(* IEC 61131-3 sources: PortalRobot/Portal_robot/Device/application (part 4) *)

(* ---- PLC_PRG.RunSafety.st ---- *)
METHOD PRIVATE RunSafety

// --- BEGIN IMPLEMENTATION ---

FOR uiTwin := 1 TO 2 DO
	axTwinSafetyBusy[uiTwin] := (GVL_TWO_PALLET.uiMode = 1) AND (GVL_TWO_PALLET.astStatus[uiTwin].xBusy
		OR (GVL_TWO_PALLET.astInput[uiTwin].xAxisBound AND NOT GVL_TWO_PALLET.astInput[uiTwin].xStandstill));
END_FOR;
FOR uiMachine := UINT#1 TO UINT#4 DO
	axButtonStationInput[uiMachine] := GVL_CELL_SAFETY_IO.axDoorUnlockButtonInput[uiMachine]
		OR ((GVL_CELL_SETTINGS.eTestEnvironment = E_CELL_TEST_ENVIRONMENT.SIMULATION)
			AND GVL_CELL_SAFETY_IO.axSimDoorUnlockButtonInput[uiMachine]);
	axButtonStationEmergencyStopInput[uiMachine] := GVL_CELL_SAFETY_IO.axEmergencyStopButtonStationInput[uiMachine]
		OR ((GVL_CELL_SETTINGS.eTestEnvironment = E_CELL_TEST_ENVIRONMENT.SIMULATION)
			AND GVL_CELL_SAFETY_IO.axSimEmergencyStopButtonStationInput[uiMachine]);
END_FOR;
CELL_SAFETY(
	axMagazineMechanismBusy := axTwinSafetyBusy,
	axDoorLockClosedInput := GVL_CELL_SAFETY_IO.axDoorLockClosedInput,
	axDoorUnlockButtonInput := axButtonStationInput,
	axEmergencyStopButtonStationInput := axButtonStationEmergencyStopInput,
	axEmergencyStopCabinetInput := GVL_CELL_SAFETY_IO.axEmergencyStopCabinetInput,
	xEmergencyStopMpgInput := GVL_CELL_SAFETY_IO.xEmergencyStopMpgInput,
	xPhaseRelayOkInput := GVL_CELL_SAFETY_IO.xPhaseRelayOkInput,
	xPressureRelayOkInput := GVL_CELL_SAFETY_IO.xPressureRelayOkInput,
	xSafetyRelayOkInput := GVL_CELL_SAFETY_IO.xSafetyRelayOkInput,
	xCellStartButtonInput := GVL_CELL_SAFETY_IO.xCellStartButtonInput,
	xCellStopButtonInput := GVL_CELL_SAFETY_IO.xCellStopButtonInput,
	xCellResetButtonInput := GVL_CELL_SAFETY_IO.xCellResetButtonInput,
	xMpgAxisXInput := GVL_CELL_SAFETY_IO.xMpgAxisXInput,
	xMpgAxisYInput := GVL_CELL_SAFETY_IO.xMpgAxisYInput,
	xMpgAxisZInput := GVL_CELL_SAFETY_IO.xMpgAxisZInput,
	xMpgMultiplier1Input := GVL_CELL_SAFETY_IO.xMpgMultiplier1Input,
	xMpgMultiplier10Input := GVL_CELL_SAFETY_IO.xMpgMultiplier10Input,
	xMpgMultiplier100Input := GVL_CELL_SAFETY_IO.xMpgMultiplier100Input,
	xSafetyRelayReset := GVL_HMI.xSafetyRelayReset,
	astMagazineStatus := GVL_MAGAZINE.astStatus,
	FaultRequest := stSafetyFaultRequest
);

GVL_CELL_SAFETY_IO.axDoorUnlockOutput := CELL_SAFETY.axDoorUnlockOutput;
GVL_CELL_SAFETY_IO.axDoorButtonLampOutput := CELL_SAFETY.axDoorButtonLampOutput;
GVL_CELL_SAFETY_IO.xSafetyRelayResetOutput := CELL_SAFETY.xSafetyRelayResetOutput;

// Физические Старт/Стоп/Сброс — равноправные дубли HMI-команд, но только по фронту.
GVL_CELL_CONTROL.xEnable := GVL_CELL_CONTROL.xEnable OR CELL_SAFETY.xCellEnablePulse;
GVL_CELL_CONTROL.xDisable := GVL_CELL_CONTROL.xDisable OR CELL_SAFETY.xCellDisablePulse;
GVL_CELL_CONTROL.xReset := GVL_CELL_CONTROL.xReset OR CELL_SAFETY.xCellResetPulse;

// Ручное I/O владеет механизмами. Физический Start также не возобновляет
// прерванный автомат; выход из этого режима сам по себе ничего не запускает.
IF xIoManualActive THEN
	GVL_CELL_CONTROL.xStart := FALSE;
	GVL_CELL_CONTROL.xEnable := FALSE;
	GVL_CELL_CONTROL.xStop := TRUE;
END_IF;

CONTROLLER_DIAGNOSTICS(
    Request := GVL_HMI.stControllerWebRequest,
    udiNowMs := udiHmiCommandNowMs,
    xReset := GVL_CELL_CONTROL.xReset,
    xResetWarnings := GVL_ALARM.Command.xResetWarnings
);
GVL_HMI.stControllerWebStatus := CONTROLLER_DIAGNOSTICS.Status;
GVL_CELL_CONTROL.xGlobalError := CELL_SAFETY.Status.xGlobalError
    OR CONTROLLER_DIAGNOSTICS.Status.xGlobalStopRequired;
IF CONTROLLER_DIAGNOSTICS.Status.xAlarmActive THEN
    // Аппаратная системная авария не допускает обход через прямые ручные DO.
    xIoManualActive := FALSE;
    // Подтверждённое исчезновение причины разрешает восстановление, но не Auto.
    GVL_CELL_CONTROL.xStart := FALSE;
    GVL_CELL_CONTROL.xEnable := FALSE;
END_IF;

// HMI записывает payload, затем CommandSeq. Gateway удерживает единственного
// писателя до AckSeq. Даже запись между RunSafety и PublishHmi не теряется:
// PLC никогда не перезаписывает запрос, а обработает его в следующем скане.
uiCellModeRejectReason := UINT#0;
udiCellModeCommandSnapshot := GVL_HMI.udiCellModeCommandSeq;
IF (udiCellModeCommandSnapshot <> UDINT#0)
AND (udiCellModeCommandSnapshot <> GVL_HMI.udiCellModeAckSeq) THEN
	IF GVL_HMI.xCellManualRequest
	AND GVL_CELL_MANAGER.Status.xRunning
	AND NOT GVL_CELL_CONTROL.xGlobalError THEN
		uiCellModeRejectReason := UINT#2;
	ELSIF NOT GVL_HMI.xCellManualRequest
	AND (GVL_CELL_CONTROL.xGlobalError OR GVL_HMI.xIoEmergencyStopActive
        OR CONTROLLER_DIAGNOSTICS.Status.xAlarmActive) THEN
		uiCellModeRejectReason := UINT#3;
	ELSE
		GVL_CELL_CONTROL.xManual := GVL_HMI.xCellManualRequest;
	END_IF;
	IF uiCellModeRejectReason = UINT#0 THEN
		GVL_HMI.uiCellModeResult := UINT#1;
	ELSE
		GVL_HMI.uiCellModeResult := uiCellModeRejectReason;
	END_IF;
	// Ack публикуется после фактического режима в PublishHmi, включая отказ.
END_IF;

IF GVL_CELL_CONTROL.xGlobalError OR GVL_HMI.xIoEmergencyStopActive
OR CONTROLLER_DIAGNOSTICS.Status.xAlarmActive THEN
	GVL_CELL_CONTROL.xManual := TRUE;
END_IF;

// Разрешения рассчитываются после применения режима и Safety текущего скана.
xRobotHmiPermit := GVL_CELL_CONTROL.xManual AND NOT GVL_CELL_MANAGER.Status.xRunning
    AND NOT xIoManualActive
    AND NOT GVL_HMI.xIoEmergencyStopActive;
xRobotAutoPowerOff := NOT GVL_CELL_CONTROL.xManual
	AND (GVL_ROBOT.Status.xError
		OR GVL_AXIS.arrAxis[1].Status.xError
		OR GVL_AXIS.arrAxis[2].Status.xError
		OR GVL_AXIS.arrAxis[3].Status.xError
		OR GVL_AXIS_GROUP.AxisGroup.Status.xLocalError
		OR GVL_AXIS_GROUP.AxisGroup.Status.xLogicalError
		OR GVL_AXIS_GROUP.AxisGroup.Status.xGroupError);

(* ---- PLC_PRG.RunSignalTower.st ---- *)
METHOD PRIVATE RunSignalTower
VAR
	xBlink : BOOL;
END_VAR

// --- BEGIN IMPLEMENTATION ---

fbAlarmHorn(astSource := astAlarmSource, tDuration := GVL_CELL_SETTINGS.tAlarmHornDuration);
GVL_CELL_SAFETY_IO.xAlarmHornOutput := fbAlarmHorn.xSound;

// Приоритет: авария > предупреждение > работа > готовность > остановлена/не готова.
// Вызывать после RunAlarms: используются актуальные сводные состояния этого скана.
IF GVL_ALARM.Status.xAlarmActive THEN
	usiSignalTowerMode := USINT#4;
ELSIF GVL_ALARM.Status.xWarningActive THEN
	usiSignalTowerMode := USINT#3;
ELSIF GVL_CELL_MANAGER.Status.xRunning THEN
	usiSignalTowerMode := USINT#1;
ELSIF GVL_CELL_MANAGER.Status.xReadyToStart THEN
	usiSignalTowerMode := USINT#2;
ELSE
	usiSignalTowerMode := USINT#5;
END_IF;

xBlink := (usiSignalTowerMode = USINT#2) OR (usiSignalTowerMode = USINT#4);
tonSignalTowerBlink(
	IN := xBlink AND (usiSignalTowerMode = usiSignalTowerPreviousMode) AND NOT tonSignalTowerBlink.Q,
	PT := T#500MS
);
// Каждый новый режим начинается со включённой секции, без ожидания таймера.
IF (usiSignalTowerMode <> usiSignalTowerPreviousMode) OR NOT xBlink THEN
	xSignalTowerBlinkOn := TRUE;
ELSIF tonSignalTowerBlink.Q THEN
	xSignalTowerBlinkOn := NOT xSignalTowerBlinkOn;
END_IF;
usiSignalTowerPreviousMode := usiSignalTowerMode;

GVL_CELL_SAFETY_IO.xSignalTowerRedOutput := (usiSignalTowerMode = USINT#5)
	OR ((usiSignalTowerMode = USINT#4) AND xSignalTowerBlinkOn);
GVL_CELL_SAFETY_IO.xSignalTowerAmberOutput := usiSignalTowerMode = USINT#3;
GVL_CELL_SAFETY_IO.xSignalTowerGreenOutput := (usiSignalTowerMode = USINT#1)
	OR ((usiSignalTowerMode = USINT#2) AND xSignalTowerBlinkOn);

(* ---- PLC_PRG.RunStatistics.st ---- *)
METHOD PRIVATE RunStatistics

// --- BEGIN IMPLEMENTATION ---

STATISTIC_MAIN(
    xStart := GVL_CELL_MANAGER.Status.xRunning,
    uiSimulationTimeFactor := GVL_CELL_SETTINGS.uiSimulationTimeFactorApplied,
    eActiveAction := GVL_ROBOT.Diag.eActiveAction,
    eActivePoint := GVL_ROBOT.Diag.eActivePoint,
    xBusyMagazine := GVL_MAGAZINE.astStatus[1].xBusy OR GVL_MAGAZINE.astStatus[2].xBusy,
    xBusyMachine_1 := GVL_MACHINE.Status[1].xBusy,
    xBusyMachine_2 := GVL_MACHINE.Status[2].xBusy,
    xBusyMachine_3 := GVL_MACHINE.Status[3].xBusy,
    xCycleActiveMachine_1 := GVL_MACHINE.Status[1].stIo.xCycleActive,
    xCycleActiveMachine_2 := GVL_MACHINE.Status[2].stIo.xCycleActive,
    xCycleActiveMachine_3 := GVL_MACHINE.Status[3].stIo.xCycleActive,
    xBusyRobot := GVL_ROBOT.Status.xBusy,
    udiNowMs := TIME_TO_UDINT(TIME())
);

IF STATISTIC_MAIN.xUpdated THEN
    GVL_STATISTIC.stStatistic := STATISTIC_MAIN.stStatistic;
END_IF;

(* ---- PLC_PRG.RunTestControl.st ---- *)
METHOD PRIVATE RunTestControl

// --- BEGIN IMPLEMENTATION ---

// Test environment is independent from the robot control interface.
rtTestEnvironmentApply(CLK := GVL_HMI.xTestEnvironmentApply);
rtTestSpeedProfileApply(CLK := GVL_HMI.xTestSpeedProfileApply);
rtTestScenarioApply(CLK := GVL_HMI.xTestScenarioApply);
xTestInitializePulse := FALSE;
xTestAbortActive := GVL_HMI.xTestAbort
	AND GVL_HMI.xTestSessionActive
	AND (GVL_CELL_SETTINGS.eTestEnvironment = E_CELL_TEST_ENVIRONMENT.SIMULATION);

xTestStable := NOT GVL_CELL_MANAGER.Status.xRunning
	AND NOT GVL_ROBOT.Status.xBusy
	AND NOT GVL_MAGAZINE.astStatus[1].xBusy
	AND NOT GVL_MAGAZINE.astStatus[2].xBusy
	AND NOT GVL_TWO_PALLET.astStatus[1].xBusy
	AND NOT GVL_TWO_PALLET.astStatus[2].xBusy
	AND NOT GVL_GEOMETRY_CONTROL.astStatus[1].xDriveRunning
	AND NOT GVL_GEOMETRY_CONTROL.astStatus[2].xDriveRunning
	AND NOT GVL_GEOMETRY_CONTROL.astStatus[1].xResetBusy
	AND NOT GVL_GEOMETRY_CONTROL.astStatus[2].xResetBusy
	AND NOT GVL_GEOMETRY_CONTROL.astStatus[1].xReserved
	AND NOT GVL_GEOMETRY_CONTROL.astStatus[2].xReserved
	AND NOT xMotionBusy
	AND NOT SIMULATION_DYNAMICS.xBusy;
FOR uiTestIndex := UINT#1 TO UINT#3 DO
	xTestStable := xTestStable
		AND NOT GVL_MACHINE.Status[uiTestIndex].xBusy
		AND NOT GVL_MACHINE.Status[uiTestIndex].xProcessing;
END_FOR;

GVL_HMI.xTestEnvironmentChangeAllowed := xTestStable
	AND NOT GVL_TWO_PALLET.astInput[1].xPowered
	AND NOT GVL_TWO_PALLET.astInput[2].xPowered;
GVL_HMI.xTestScenarioApplyAllowed := xTestStable
	AND ((GVL_TWO_PALLET.uiMode = 0)
		OR ((GVL_TWO_PALLET.uiMode = 1)
			AND (GVL_CELL_SETTINGS.eTestEnvironment = E_CELL_TEST_ENVIRONMENT.SIMULATION)
			AND NOT GVL_HMI.xModbusMode
			AND GVL_TWO_PALLET.astStatus[1].xConfirmed
			AND GVL_TWO_PALLET.astStatus[2].xConfirmed
			AND (GVL_TWO_PALLET.astStatus[1].uiRobotPallet >= UINT#1)
			AND (GVL_TWO_PALLET.astStatus[1].uiRobotPallet <= UINT#2)
			AND (GVL_TWO_PALLET.astStatus[2].uiRobotPallet >= UINT#1)
			AND (GVL_TWO_PALLET.astStatus[2].uiRobotPallet <= UINT#2)
			AND GVL_TWO_PALLET.astInput[1].xStandstill
			AND GVL_TWO_PALLET.astInput[2].xStandstill))
	AND GVL_HMI.xTestSessionActive
	AND (GVL_CELL_SETTINGS.eTestEnvironment <> E_CELL_TEST_ENVIRONMENT.NORMAL)
	AND ((GVL_CELL_SETTINGS.eTestEnvironment <> E_CELL_TEST_ENVIRONMENT.SIMULATION)
		OR NOT GVL_ROBOT_MODBUS.xModeActive
		OR GVL_ROBOT_MODBUS.Status.xSimulatorActive);
// Старые OPC UA поля сохранены для совместимости; физический ключ исключён.
GVL_HMI.xSc500BenchKeyActive := FALSE;

IF rtTestEnvironmentApply.Q THEN
	GVL_HMI.uiTestRejectReason := UINT#0;
	IF NOT GVL_HMI.xTestEnvironmentChangeAllowed THEN
		GVL_HMI.uiTestRejectReason := UINT#1; // equipment is not idle
	ELSIF GVL_HMI.uiTestEnvironmentRequest > UINT#2 THEN
		GVL_HMI.uiTestRejectReason := UINT#2; // invalid environment
	ELSIF (GVL_HMI.uiTestEnvironmentRequest = UINT#2)
	AND NOT GVL_ROBOT_MODBUS.xModeActive THEN
		GVL_HMI.uiTestRejectReason := UINT#3; // bench requires Modbus
	ELSIF (GVL_HMI.uiTestEnvironmentRequest = UINT#1)
	AND GVL_ROBOT_MODBUS.xModeActive
	AND NOT GVL_ROBOT_MODBUS.Status.xSimulatorActive THEN
		GVL_HMI.uiTestRejectReason := UINT#4; // Python simulator marker missing
	ELSE
		CASE GVL_HMI.uiTestEnvironmentRequest OF
			UINT#0: GVL_CELL_SETTINGS.eTestEnvironment := E_CELL_TEST_ENVIRONMENT.NORMAL;
			UINT#1: GVL_CELL_SETTINGS.eTestEnvironment := E_CELL_TEST_ENVIRONMENT.SIMULATION;
			UINT#2: GVL_CELL_SETTINGS.eTestEnvironment := E_CELL_TEST_ENVIRONMENT.SC500_BENCH;
		END_CASE;
		IF GVL_CELL_SETTINGS.eTestEnvironment = E_CELL_TEST_ENVIRONMENT.NORMAL THEN
			GVL_CELL_SETTINGS.xErrorSimulationEnabled := FALSE;
		END_IF;
		GVL_CELL_SETTINGS.eTestSpeedProfile := E_TEST_SPEED_PROFILE.REALTIME;
	END_IF;
END_IF;

IF rtTestSpeedProfileApply.Q THEN
	GVL_HMI.uiTestRejectReason := UINT#0;
	IF (GVL_HMI.uiTestSpeedProfileRequest <= UINT#1)
	AND (GVL_CELL_SETTINGS.eTestEnvironment = E_CELL_TEST_ENVIRONMENT.SIMULATION) THEN
		IF GVL_HMI.uiTestSpeedProfileRequest = UINT#1 THEN
			GVL_CELL_SETTINGS.eTestSpeedProfile := E_TEST_SPEED_PROFILE.FAST;
			// В Modbus профиль по-прежнему владеет коэффициентом внешней модели.
			// В SoftMotion коэффициент задаёт ползунок, а применение выполняется
			// отдельной транзакцией только на границе следующего теста.
			IF GVL_ROBOT_MODBUS.xModeActive THEN
				GVL_CELL_SETTINGS.uiSimulationTimeFactor := UINT#250;
			END_IF;
		ELSE
			GVL_CELL_SETTINGS.eTestSpeedProfile := E_TEST_SPEED_PROFILE.REALTIME;
			IF GVL_ROBOT_MODBUS.xModeActive THEN
				GVL_CELL_SETTINGS.uiSimulationTimeFactor := UINT#1;
			END_IF;
		END_IF;
		GVL_HMI.uiSimulationTimeFactor := GVL_CELL_SETTINGS.uiSimulationTimeFactor;
	ELSE
		GVL_HMI.uiTestRejectReason := UINT#5; // speed profile is simulation-only
	END_IF;
END_IF;

IF rtTestScenarioApply.Q THEN
	GVL_HMI.uiTestScenarioResult := UINT#0;
	uiTestSlotCount := UINT#120;
	IF GVL_TWO_PALLET.uiMode = UINT#1 THEN uiTestSlotCount := UINT#96; END_IF;
	xTestScenarioValid := (GVL_HMI.stTestScenario.uiSchemaVersion = UINT#3)
		AND (GVL_HMI.stTestScenario.uiMagazineMode = GVL_TWO_PALLET.uiMode)
		AND (GVL_HMI.stTestScenario.udiLoadSeq <> UDINT#0)
		AND (GVL_HMI.stTestScenario.uiTypeCount >= UINT#1)
		AND (GVL_HMI.stTestScenario.uiTypeCount <= UINT#3);
	FOR uiTestIndex := UINT#1 TO UINT#3 DO
		xTestScenarioValid := xTestScenarioValid
			AND (GVL_HMI.stTestScenario.auiMachineState[uiTestIndex] <= UINT#3)
			AND (GVL_HMI.stTestScenario.auiMachineType[uiTestIndex] >= UINT#1)
			AND (GVL_HMI.stTestScenario.auiMachineType[uiTestIndex]
				<= GVL_HMI.stTestScenario.uiTypeCount);
	END_FOR;
	FOR uiTestIndex := UINT#1 TO uiTestSlotCount DO
		xTestScenarioValid := xTestScenarioValid
			AND (GVL_HMI.stTestScenario.auiSlotType[uiTestIndex] >= UINT#1)
			AND (GVL_HMI.stTestScenario.auiSlotType[uiTestIndex]
				<= GVL_HMI.stTestScenario.uiTypeCount);
		FOR uiTestMagazine := UINT#1 TO UINT#2 DO
			xTestScenarioValid := xTestScenarioValid
				AND (GVL_HMI.stTestScenario.aauiSlotContent[uiTestMagazine, uiTestIndex] <= UINT#2)
				AND (GVL_HMI.stTestScenario.aauiOperatorSlotContent[uiTestMagazine, uiTestIndex] <= UINT#2);
		END_FOR;
	END_FOR;
	FOR uiTestType := UINT#1 TO MIN(UINT#3, GVL_HMI.stTestScenario.uiTypeCount) DO
		xTestTypeHasMachine := FALSE;
		xTestTypeHasSlot := FALSE;
		FOR uiTestIndex := UINT#1 TO UINT#3 DO
			xTestTypeHasMachine := xTestTypeHasMachine OR (GVL_HMI.stTestScenario.auiMachineType[uiTestIndex] = uiTestType);
		END_FOR;
		FOR uiTestIndex := UINT#1 TO uiTestSlotCount DO
			xTestTypeHasSlot := xTestTypeHasSlot OR (GVL_HMI.stTestScenario.auiSlotType[uiTestIndex] = uiTestType);
		END_FOR;
		xTestScenarioValid := xTestScenarioValid AND xTestTypeHasMachine AND xTestTypeHasSlot;
	END_FOR;
	uiTestFaultOwnerCount := UINT#0;
	IF GVL_HMI.stTestScenario.dwCellFaultMask <> DWORD#0 THEN
		uiTestFaultOwnerCount := uiTestFaultOwnerCount + UINT#1;
	END_IF;
	IF GVL_HMI.stTestScenario.dwRobotFaultMask <> DWORD#0 THEN
		uiTestFaultOwnerCount := uiTestFaultOwnerCount + UINT#1;
	END_IF;
	FOR uiTestMagazine := UINT#1 TO UINT#2 DO
		IF GVL_HMI.stTestScenario.adwMagazineFaultMask[uiTestMagazine] <> DWORD#0 THEN
			uiTestFaultOwnerCount := uiTestFaultOwnerCount + UINT#1;
		END_IF;
		xTestScenarioValid := xTestScenarioValid
			AND (GVL_HMI.stTestScenario.adwMagazineFaultMask[uiTestMagazine] <= DWORD#16#0000_003F);
	END_FOR;
	FOR uiTestIndex := UINT#1 TO UINT#3 DO
		IF GVL_HMI.stTestScenario.adwMachineFaultMask[uiTestIndex] <> DWORD#0 THEN
			uiTestFaultOwnerCount := uiTestFaultOwnerCount + UINT#1;
		END_IF;
		xTestScenarioValid := xTestScenarioValid
			AND (GVL_HMI.stTestScenario.adwMachineFaultMask[uiTestIndex] <= DWORD#16#0000_07FF);
	END_FOR;
	xTestScenarioValid := xTestScenarioValid
		AND (uiTestFaultOwnerCount <= UINT#1)
		AND (GVL_HMI.stTestScenario.dwCellFaultMask <= DWORD#16#0000_0001)
		AND (GVL_HMI.stTestScenario.dwRobotFaultMask <= DWORD#16#0000_01FF)
		AND (GVL_HMI.stTestScenario.auiGripperContent[1] <= UINT#1)
		AND ((GVL_HMI.stTestScenario.auiGripperContent[1] = UINT#0)
			= (GVL_HMI.stTestScenario.auiGripperType[1] = UINT#0))
		AND (GVL_HMI.stTestScenario.auiGripperType[1]
			<= GVL_HMI.stTestScenario.uiTypeCount)
		AND ((GVL_HMI.stTestScenario.auiGripperContent[2] = UINT#0)
			OR (GVL_HMI.stTestScenario.auiGripperContent[2] = UINT#2))
		AND ((GVL_HMI.stTestScenario.auiGripperContent[2] = UINT#0)
			= (GVL_HMI.stTestScenario.auiGripperType[2] = UINT#0))
		AND (GVL_HMI.stTestScenario.auiGripperType[2]
			<= GVL_HMI.stTestScenario.uiTypeCount);

	IF GVL_HMI.stTestScenario.axGeometryEnabled[1] OR GVL_HMI.stTestScenario.axGeometryEnabled[2]
		OR GVL_HMI.stTestScenario.axGeometryCall[1] OR GVL_HMI.stTestScenario.axGeometryCall[2]
		OR GVL_HMI.stTestScenario.axGeometryCall[3] THEN
		xTestScenarioValid := xTestScenarioValid
			AND (GVL_CELL_SETTINGS.eTestEnvironment = E_CELL_TEST_ENVIRONMENT.SIMULATION)
			AND NOT GVL_HMI.xModbusMode;
	END_IF;
	IF NOT GVL_HMI.xTestScenarioApplyAllowed THEN
		GVL_HMI.uiTestScenarioResult := UINT#1;
	ELSIF NOT xTestScenarioValid OR (GVL_HMI.stTestScenario.uiOrientation > UINT#1) THEN
		GVL_HMI.uiTestScenarioResult := UINT#2;
	ELSE
		FOR uiTestMagazine := UINT#1 TO UINT#2 DO
			uiTestPallet := GVL_TWO_PALLET.astStatus[uiTestMagazine].uiRobotPallet;
			uiTestOtherPallet := UINT#3 - uiTestPallet;
			FOR uiTestIndex := UINT#1 TO UINT#120 DO
				GVL_DETAIL.astMagazine[uiTestMagazine].aSlots[uiTestIndex].xInPosition := FALSE;
				GVL_DETAIL.astMagazine[uiTestMagazine].aSlots[uiTestIndex].eDetailType := E_DETAIL_TYPE.NONE;
				GVL_DETAIL.astMagazine[uiTestMagazine].aSlots[uiTestIndex].uiProductType := UINT#0;
				IF uiTestIndex <= uiTestSlotCount THEN
					GVL_DETAIL.astMagazine[uiTestMagazine].aSlots[uiTestIndex].xInPosition :=
						GVL_HMI.stTestScenario.aauiSlotContent[uiTestMagazine, uiTestIndex] <> UINT#0;
					CASE GVL_HMI.stTestScenario.aauiSlotContent[uiTestMagazine, uiTestIndex] OF
						UINT#1: GVL_DETAIL.astMagazine[uiTestMagazine].aSlots[uiTestIndex].eDetailType := E_DETAIL_TYPE.BLANK;
						UINT#2: GVL_DETAIL.astMagazine[uiTestMagazine].aSlots[uiTestIndex].eDetailType := E_DETAIL_TYPE.DETAIL;
					END_CASE;
					IF GVL_DETAIL.astMagazine[uiTestMagazine].aSlots[uiTestIndex].xInPosition THEN
						GVL_DETAIL.astMagazine[uiTestMagazine].aSlots[uiTestIndex].uiProductType := GVL_HMI.stTestScenario.auiSlotType[uiTestIndex];
					END_IF;
				END_IF;
				IF GVL_TWO_PALLET.uiMode = UINT#1 THEN
					GVL_TWO_PALLET.astStore[uiTestMagazine].astPallet[uiTestPallet].aSlots[uiTestIndex] := GVL_DETAIL.astMagazine[uiTestMagazine].aSlots[uiTestIndex];
					GVL_TWO_PALLET.astStore[uiTestMagazine].astPallet[uiTestOtherPallet].aSlots[uiTestIndex].xInPosition := FALSE;
					GVL_TWO_PALLET.astStore[uiTestMagazine].astPallet[uiTestOtherPallet].aSlots[uiTestIndex].eDetailType := E_DETAIL_TYPE.NONE;
					GVL_TWO_PALLET.astStore[uiTestMagazine].astPallet[uiTestOtherPallet].aSlots[uiTestIndex].uiProductType := UINT#0;
					IF uiTestIndex <= uiTestSlotCount THEN
						GVL_TWO_PALLET.astStore[uiTestMagazine].astPallet[uiTestOtherPallet].aSlots[uiTestIndex].xInPosition := GVL_HMI.stTestScenario.aauiOperatorSlotContent[uiTestMagazine, uiTestIndex] <> UINT#0;
						CASE GVL_HMI.stTestScenario.aauiOperatorSlotContent[uiTestMagazine, uiTestIndex] OF
							UINT#1: GVL_TWO_PALLET.astStore[uiTestMagazine].astPallet[uiTestOtherPallet].aSlots[uiTestIndex].eDetailType := E_DETAIL_TYPE.BLANK;
							UINT#2: GVL_TWO_PALLET.astStore[uiTestMagazine].astPallet[uiTestOtherPallet].aSlots[uiTestIndex].eDetailType := E_DETAIL_TYPE.DETAIL;
						END_CASE;
						IF GVL_HMI.stTestScenario.aauiOperatorSlotContent[uiTestMagazine, uiTestIndex] <> UINT#0 THEN
							GVL_TWO_PALLET.astStore[uiTestMagazine].astPallet[uiTestOtherPallet].aSlots[uiTestIndex].uiProductType := GVL_HMI.stTestScenario.auiSlotType[uiTestIndex];
						END_IF;
					END_IF;
				END_IF;
			END_FOR;
			IF GVL_TWO_PALLET.uiMode = UINT#1 THEN
				GVL_TWO_PALLET.astStore[uiTestMagazine].axLoaded[uiTestPallet] := FALSE;
				GVL_TWO_PALLET.astStore[uiTestMagazine].axLoaded[uiTestOtherPallet] := GVL_HMI.stTestScenario.axOperatorLoaded[uiTestMagazine];
				GVL_TWO_PALLET.axSimulationAutoSwapEnabled[uiTestMagazine] := GVL_HMI.stTestScenario.axAutoSwap[uiTestMagazine];
			ELSE
				GVL_TWO_PALLET.astStatic[uiTestMagazine] := GVL_DETAIL.astMagazine[uiTestMagazine];
			END_IF;
			adwTestMagazineFaultMask[uiTestMagazine] := GVL_HMI.stTestScenario.adwMagazineFaultMask[uiTestMagazine];
		END_FOR;
		// Начальные инъекции: маски переводятся в существующий диагностический
		// контракт, а не обходят владельцев ошибок.
		axHmiInternalPulse[13] :=
			(GVL_HMI.stTestScenario.dwCellFaultMask AND DWORD#16#0000_0001) <> DWORD#0;
		axHmiInternalPulse[12] :=
			(GVL_HMI.stTestScenario.dwRobotFaultMask AND DWORD#16#0000_0001) <> DWORD#0;
		GVL_HMI.xSimGripper1Fault :=
			(GVL_HMI.stTestScenario.dwRobotFaultMask AND DWORD#16#0000_0002) <> DWORD#0;
		GVL_HMI.xSimGripper2Fault :=
			(GVL_HMI.stTestScenario.dwRobotFaultMask AND DWORD#16#0000_0004) <> DWORD#0;
		GVL_HMI.xSimGripperRotationFault :=
			(GVL_HMI.stTestScenario.dwRobotFaultMask AND DWORD#16#0000_0008) <> DWORD#0;
		GVL_HMI.xSimGripperGlobalFault :=
			(GVL_HMI.stTestScenario.dwRobotFaultMask AND DWORD#16#0000_0010) <> DWORD#0;
		axHmiInternalPulse[14] :=
			(GVL_HMI.stTestScenario.dwRobotFaultMask AND DWORD#16#0000_0020) <> DWORD#0;
		axHmiInternalPulse[15] :=
			(GVL_HMI.stTestScenario.dwRobotFaultMask AND DWORD#16#0000_0040) <> DWORD#0;
		axHmiInternalPulse[16] :=
			(GVL_HMI.stTestScenario.dwRobotFaultMask AND DWORD#16#0000_0080) <> DWORD#0;
		axHmiInternalPulse[17] :=
			(GVL_HMI.stTestScenario.dwRobotFaultMask AND DWORD#16#0000_0100) <> DWORD#0;
		axHmiInternalPulse[18] :=
			(GVL_HMI.stTestScenario.adwMagazineFaultMask[1] AND DWORD#16#0000_0001) <> DWORD#0;
		axHmiInternalPulse[19] :=
			(GVL_HMI.stTestScenario.adwMagazineFaultMask[1] AND DWORD#16#0000_0002) <> DWORD#0;
		axHmiInternalPulse[20] :=
			(GVL_HMI.stTestScenario.adwMagazineFaultMask[1] AND DWORD#16#0000_0004) <> DWORD#0;
		axHmiInternalPulse[21] :=
			(GVL_HMI.stTestScenario.adwMagazineFaultMask[1] AND DWORD#16#0000_0008) <> DWORD#0;
		axHmiInternalPulse[22] :=
			(GVL_HMI.stTestScenario.adwMagazineFaultMask[1] AND DWORD#16#0000_0010) <> DWORD#0;
		axHmiInternalPulse[23] :=
			(GVL_HMI.stTestScenario.adwMagazineFaultMask[1] AND DWORD#16#0000_0020) <> DWORD#0;
		FOR uiTestIndex := UINT#1 TO UINT#3 DO
			GVL_HMI.axMachineSimAlarm[uiTestIndex] :=
				(GVL_HMI.stTestScenario.adwMachineFaultMask[uiTestIndex] AND DWORD#16#0000_0001) <> DWORD#0;
			GVL_HMI.axMachineSimDoorFault[uiTestIndex] :=
				(GVL_HMI.stTestScenario.adwMachineFaultMask[uiTestIndex] AND DWORD#16#0000_0002) <> DWORD#0;
			GVL_HMI.axMachineSimChuckFault[uiTestIndex] :=
				(GVL_HMI.stTestScenario.adwMachineFaultMask[uiTestIndex] AND DWORD#16#0000_0004) <> DWORD#0;
			GVL_HMI.axMachineTimeoutRobotMove[uiTestIndex] :=
				(GVL_HMI.stTestScenario.adwMachineFaultMask[uiTestIndex] AND DWORD#16#0000_0008) <> DWORD#0;
			GVL_HMI.axMachineTimeoutRobotAction[uiTestIndex] :=
				(GVL_HMI.stTestScenario.adwMachineFaultMask[uiTestIndex] AND DWORD#16#0000_0010) <> DWORD#0;
			GVL_HMI.axMachineTimeoutRobotRelease[uiTestIndex] :=
				(GVL_HMI.stTestScenario.adwMachineFaultMask[uiTestIndex] AND DWORD#16#0000_0020) <> DWORD#0;
			GVL_HMI.axMachineTimeoutDoorOpen[uiTestIndex] :=
				(GVL_HMI.stTestScenario.adwMachineFaultMask[uiTestIndex] AND DWORD#16#0000_0040) <> DWORD#0;
			GVL_HMI.axMachineTimeoutDoorClose[uiTestIndex] :=
				(GVL_HMI.stTestScenario.adwMachineFaultMask[uiTestIndex] AND DWORD#16#0000_0080) <> DWORD#0;
			GVL_HMI.axMachineTimeoutChuckOpen[uiTestIndex] :=
				(GVL_HMI.stTestScenario.adwMachineFaultMask[uiTestIndex] AND DWORD#16#0000_0100) <> DWORD#0;
			GVL_HMI.axMachineTimeoutChuckClose[uiTestIndex] :=
				(GVL_HMI.stTestScenario.adwMachineFaultMask[uiTestIndex] AND DWORD#16#0000_0200) <> DWORD#0;
			GVL_HMI.axMachineTimeoutCycleStart[uiTestIndex] :=
				(GVL_HMI.stTestScenario.adwMachineFaultMask[uiTestIndex] AND DWORD#16#0000_0400) <> DWORD#0;
		END_FOR;
		GVL_HMI.xErrorSimulationEnable :=
			(GVL_HMI.stTestScenario.dwCellFaultMask <> DWORD#0)
			OR (GVL_HMI.stTestScenario.dwRobotFaultMask <> DWORD#0)
			OR (GVL_HMI.stTestScenario.adwMagazineFaultMask[1] <> DWORD#0)
			OR (GVL_HMI.stTestScenario.adwMagazineFaultMask[2] <> DWORD#0)
			OR (GVL_HMI.stTestScenario.adwMachineFaultMask[1] <> DWORD#0)
			OR (GVL_HMI.stTestScenario.adwMachineFaultMask[2] <> DWORD#0)
			OR (GVL_HMI.stTestScenario.adwMachineFaultMask[3] <> DWORD#0);
		IF GVL_CELL_SETTINGS.eTestEnvironment = E_CELL_TEST_ENVIRONMENT.SIMULATION THEN
			IF NOT xTestGeometrySettingsSaved THEN
				xTestSavedGeometryAuto := Persistent_Value.xAutoEnabled;
				xTestSavedGeometryWait := Persistent_Value.xWaitWhenOccupied;
				xTestGeometrySettingsSaved := TRUE;
			END_IF;
			Persistent_Value.xAutoEnabled := FALSE;
			Persistent_Value.xWaitWhenOccupied := GVL_HMI.stTestScenario.xGeometryWaitWhenOccupied;
		END_IF;
		xTestInitializePulse := TRUE;
	END_IF;
	// Ack подтверждает обработку конкретного LoadSeq даже при отклонении.
	GVL_HMI.udiTestScenarioAckSeq := GVL_HMI.stTestScenario.udiLoadSeq;
END_IF;

GVL_HMI.uiTestEnvironmentApplied := TO_UINT(GVL_CELL_SETTINGS.eTestEnvironment);
GVL_HMI.uiTestSpeedProfileApplied := TO_UINT(GVL_CELL_SETTINGS.eTestSpeedProfile);
GVL_HMI.xSc500BenchKeyLost := FALSE;
IF GVL_CELL_SETTINGS.eTestEnvironment = E_CELL_TEST_ENVIRONMENT.SIMULATION THEN
	IF GVL_HMI.xTestSessionActive THEN
		GVL_CELL_SETTINGS.xSimulationAccelerationEnable :=
			GVL_CELL_SETTINGS.eTestSpeedProfile = E_TEST_SPEED_PROFILE.FAST;
		// Профиль владеет включением ускоренных таймеров, а сам коэффициент
		// разрешено менять с HMI прямо во время тестового движения.
		GVL_HMI.xSimulationAccelerationEnable := GVL_CELL_SETTINGS.xSimulationAccelerationEnable;
	END_IF;
ELSE
	GVL_CELL_SETTINGS.xSimulationAccelerationEnable := FALSE;
	GVL_HMI.xSimulationAccelerationEnable := FALSE;
END_IF;

// Restore the operator policy even if the runner crashes and gateway releases the session.
IF xTestGeometrySettingsSaved AND NOT GVL_HMI.xTestSessionActive THEN
	Persistent_Value.xAutoEnabled := xTestSavedGeometryAuto;
	Persistent_Value.xWaitWhenOccupied := xTestSavedGeometryWait;
	xTestGeometrySettingsSaved := FALSE;
END_IF;

(* ---- PLC_PRG.RunTwoPallet.st ---- *)
METHOD PRIVATE RunTwoPallet

// --- BEGIN IMPLEMENTATION ---

GVL_TWO_PALLET.xModeChanged := FALSE;
IF NOT xTwinSimulationInitialized THEN
	FOR uiTwin := 1 TO 2 DO
		// Числа используются только для виртуальных SoftMotion-осей.
		GVL_TWO_PALLET.astSimulationConfig[uiTwin].xConfigured := TRUE;
		GVL_TWO_PALLET.astSimulationConfig[uiTwin].xP1LockOut := TRUE;
		GVL_TWO_PALLET.axSimulationAutoSwapEnabled[uiTwin] := TRUE;
		GVL_TWO_PALLET.astSimulationConfig[uiTwin].lrExchange := 0.0;
		GVL_TWO_PALLET.astSimulationConfig[uiTwin].lrWorkP1 := 100.0;
		GVL_TWO_PALLET.astSimulationConfig[uiTwin].lrWorkP2 := 200.0;
		GVL_TWO_PALLET.astSimulationConfig[uiTwin].lrHome := 0.0;
		GVL_TWO_PALLET.astSimulationConfig[uiTwin].lrTolerance := 1.0;
		GVL_TWO_PALLET.astSimulationConfig[uiTwin].lrVelocity := 100.0;
		GVL_TWO_PALLET.astSimulationConfig[uiTwin].lrAcceleration := 200.0;
		GVL_TWO_PALLET.astSimulationConfig[uiTwin].lrDeceleration := 200.0;
		GVL_TWO_PALLET.astSimulationConfig[uiTwin].lrJerk := 1000.0;
		GVL_TWO_PALLET.astSimulationConfig[uiTwin].tCylinder := T#3S;
		GVL_TWO_PALLET.astSimulationConfig[uiTwin].tMove := T#20S;
		GVL_TWO_PALLET.astSimulationConfig[uiTwin].tHome := T#10S;
		GVL_TWO_PALLET.astSimulationConfig[uiTwin].tPulse := T#150MS;
	END_FOR;
	IF NOT GVL_TWO_PALLET.xAutoSwapDefaultsApplied THEN
		FOR uiTwin := 1 TO 2 DO
			GVL_TWO_PALLET.axAutoSwapEnabled[uiTwin] := TRUE;
		END_FOR;
		GVL_TWO_PALLET.xAutoSwapDefaultsApplied := TRUE;
	END_IF;
	xTwinSimulationInitialized := TRUE;
END_IF;
FOR uiTwin := 1 TO 2 DO
	GVL_TWO_PALLET.auiCommand[uiTwin] := UINT#0;
    axMagazineInventoryChanged[uiTwin] := NOT xTwinStartup OR xTestInitializePulse;
    axTwinStoreChanged[uiTwin] := NOT xTwinStartup OR xTestInitializePulse;
END_FOR;
IF NOT xTwinStartup THEN
	IF GVL_TWO_PALLET.uiMode = 0 THEN
		GVL_HMI.MagazinePitchX := Persistent_Value.lrStaticPitchX;
		GVL_HMI.MagazinePitchY := Persistent_Value.lrStaticPitchY;
	ELSE
		GVL_HMI.MagazinePitchX := Persistent_Value.lrTwinPitchX;
		GVL_HMI.MagazinePitchY := Persistent_Value.lrTwinPitchY;
	END_IF;
	FOR uiTwin := 1 TO 2 DO
		// После перезапуска содержимое сохранено, готовность загрузки подтверждается заново.
		GVL_TWO_PALLET.astStore[uiTwin].axLoaded[1] := FALSE;
		GVL_TWO_PALLET.astStore[uiTwin].axLoaded[2] := FALSE;
		axTwinStoreChanged[uiTwin] := TRUE;
		IF GVL_TWO_PALLET.uiMode = 0 THEN
			GVL_DETAIL.astMagazine[uiTwin] := GVL_TWO_PALLET.astStatic[uiTwin];
		END_IF;
	END_FOR;
	xTwinStartup := TRUE;
END_IF;
GVL_TWO_PALLET.xModeChangeAllowed := GVL_CELL_CONTROL.xManual
	AND NOT GVL_CELL_MANAGER.Status.xRunning AND NOT GVL_ROBOT.Status.xBusy AND NOT xMotionBusy
	AND xHmiConnectionAlive AND NOT GVL_HMI.xTestSessionActive AND NOT GVL_ROBOT.Status.xBlankAvailable AND NOT GVL_ROBOT.Status.xDetailAvailable
	AND (GVL_ROBOT.Status.uiMagazineContext = 0)
	AND NOT GVL_MAGAZINE.astStatus[1].xEnabled AND NOT GVL_MAGAZINE.astStatus[2].xEnabled
	AND NOT GVL_MAGAZINE.astStatus[1].xBusy AND NOT GVL_MAGAZINE.astStatus[2].xBusy
	AND NOT GVL_TWO_PALLET.astStatus[1].xBusy AND NOT GVL_TWO_PALLET.astStatus[2].xBusy
	AND NOT GVL_TWO_PALLET.astInput[1].xPowered AND NOT GVL_TWO_PALLET.astInput[2].xPowered
	AND NOT GVL_TWO_PALLET.astStatus[1].xError AND NOT GVL_TWO_PALLET.astStatus[2].xError;

udiTwinSnapshot := GVL_HMI.udiTwinCommandSeq;
uiTwinRequestResult := 0;
xTwinInventoryCommand := FALSE;
IF (udiTwinSnapshot <> 0) AND (udiTwinSnapshot <> GVL_HMI.udiTwinAckSeq) THEN
	stTwinRequest := GVL_HMI.stTwinRequest;
	uiTwinRequestResult := 2; // Условие команды не выполнено
	IF (GVL_HMI.udiHmiCommandClockMs - GVL_HMI.udiTwinIssuedAtMs) > 2000 THEN
		uiTwinRequestResult := 4;
	ELSIF (stTwinRequest.uiMagazine = 0) AND (stTwinRequest.uiCommand = 25) THEN
		IF GVL_TWO_PALLET.xModeChangeAllowed AND (stTwinRequest.uiValue <= 1) AND xHmiConnectionAlive THEN
			IF GVL_TWO_PALLET.uiMode <> stTwinRequest.uiValue THEN
				IF GVL_TWO_PALLET.uiMode = 0 THEN
					Persistent_Value.lrStaticPitchX := GVL_HMI.MagazinePitchX;
					Persistent_Value.lrStaticPitchY := GVL_HMI.MagazinePitchY;
				ELSE
					Persistent_Value.lrTwinPitchX := GVL_HMI.MagazinePitchX;
					Persistent_Value.lrTwinPitchY := GVL_HMI.MagazinePitchY;
				END_IF;
				GVL_TWO_PALLET.uiMode := stTwinRequest.uiValue;
				GVL_TWO_PALLET.xModeChanged := TRUE;
				FOR uiTwin := 1 TO 2 DO
					axMagazineInventoryChanged[uiTwin] := TRUE;
					IF GVL_TWO_PALLET.uiMode = 0 THEN GVL_DETAIL.astMagazine[uiTwin] := GVL_TWO_PALLET.astStatic[uiTwin]; END_IF;
					// Базы меняются вместе с механикой: старые координаты нельзя молча использовать.
					InvalidateMagazineCalibration(uiMagazine := uiTwin);
					axMagazinePointsReady[uiTwin] := FALSE;
				END_FOR;
				GVL_POINT.Points[E_POINT_NAME.MAGAZINE_1_DETAIL].xConfigured := FALSE;
				GVL_POINT.Points[E_POINT_NAME.MAGAZINE_2_DETAIL].xConfigured := FALSE;
				IF GVL_TWO_PALLET.uiMode = 0 THEN
					GVL_HMI.MagazinePitchX := Persistent_Value.lrStaticPitchX; GVL_HMI.MagazinePitchY := Persistent_Value.lrStaticPitchY;
				ELSE
					GVL_HMI.MagazinePitchX := Persistent_Value.lrTwinPitchX; GVL_HMI.MagazinePitchY := Persistent_Value.lrTwinPitchY;
				END_IF;
				xPointTableReady := FALSE;
			END_IF;
			uiTwinRequestResult := 1;
		END_IF;
	ELSIF (stTwinRequest.uiMagazine >= 1) AND (stTwinRequest.uiMagazine <= 2)
		AND (GVL_TWO_PALLET.uiMode = 1) THEN
		uiTwin := stTwinRequest.uiMagazine;
		IF ((stTwinRequest.uiCommand >= 1) AND (stTwinRequest.uiCommand <= 19))
			OR ((stTwinRequest.uiCommand >= 25) AND (stTwinRequest.uiCommand <= 32)) THEN
			GVL_TWO_PALLET.auiCommand[uiTwin] := stTwinRequest.uiCommand;
			GVL_TWO_PALLET.auiValue[uiTwin] := stTwinRequest.uiValue;
			GVL_TWO_PALLET.audiRevision[uiTwin] := stTwinRequest.udiRevision;
		ELSIF (stTwinRequest.uiCommand >= UINT#20)
			AND (stTwinRequest.uiCommand <= UINT#24) THEN
			xTwinInventoryCommand := TRUE; // Проверить по разрешениям текущего скана ПОСЛЕ вызова FB
		ELSIF stTwinRequest.uiCommand = UINT#33 THEN
			IF (stTwinRequest.uiValue <= UINT#1) AND xHmiConnectionAlive THEN
				IF GVL_CELL_SETTINGS.eTestEnvironment = E_CELL_TEST_ENVIRONMENT.SIMULATION THEN
					GVL_TWO_PALLET.axSimulationAutoSwapEnabled[uiTwin] := stTwinRequest.uiValue = UINT#1;
				ELSE
					GVL_TWO_PALLET.axAutoSwapEnabled[uiTwin] := stTwinRequest.uiValue = UINT#1;
				END_IF;
				uiTwinRequestResult := UINT#1;
			END_IF;
		END_IF;
	END_IF;
END_IF;

FOR uiTwin := 1 TO 2 DO
	GVL_TWO_PALLET.astActiveConfig[uiTwin] := GVL_TWO_PALLET.astConfig[uiTwin];
	IF GVL_CELL_SETTINGS.eTestEnvironment = E_CELL_TEST_ENVIRONMENT.SIMULATION THEN
		GVL_TWO_PALLET.astActiveConfig[uiTwin] := GVL_TWO_PALLET.astSimulationConfig[uiTwin];
		xTwinAutoSwapEnabled := GVL_TWO_PALLET.axSimulationAutoSwapEnabled[uiTwin];
	ELSE
		xTwinAutoSwapEnabled := GVL_TWO_PALLET.axAutoSwapEnabled[uiTwin];
	END_IF;
	// Старые RETAIN-параметры сохраняют прежнюю полярность до первой настройки
	// полных сочетаний. Нормализуем только рабочую копию, без записи в RETAIN.
	IF NOT GVL_TWO_PALLET.astActiveConfig[uiTwin].xSignalPatternsConfigured THEN
		GVL_TWO_PALLET.astActiveConfig[uiTwin].uiP1Signals := UINT#38;
		GVL_TWO_PALLET.astActiveConfig[uiTwin].uiP2Signals := UINT#26;
		IF GVL_TWO_PALLET.astActiveConfig[uiTwin].xP1LockOut THEN
			GVL_TWO_PALLET.astActiveConfig[uiTwin].uiP1Signals := UINT#26;
			GVL_TWO_PALLET.astActiveConfig[uiTwin].uiP2Signals := UINT#38;
		END_IF;
		GVL_TWO_PALLET.astActiveConfig[uiTwin].xSignalPatternsConfigured := TRUE;
	END_IF;
	// Legacy power/reset также проходит владельца механизма и его блокировки.
	IF (GVL_TWO_PALLET.auiCommand[uiTwin] = 0) AND (GVL_TWO_PALLET.uiMode = 1) THEN
		IF GVL_HMI.astMagazineCommand[uiTwin].xEnable THEN GVL_TWO_PALLET.auiCommand[uiTwin] := 1; END_IF;
		IF GVL_HMI.astMagazineCommand[uiTwin].xDisable THEN GVL_TWO_PALLET.auiCommand[uiTwin] := 3; END_IF;
		IF GVL_HMI.astMagazineCommand[uiTwin].xStop THEN GVL_TWO_PALLET.auiCommand[uiTwin] := 15; END_IF;
		IF GVL_HMI.astMagazineCommand[uiTwin].xReset
			OR (GVL_CELL_CONTROL.xReset AND GVL_TWO_PALLET.astStatus[uiTwin].xResetAllowed) THEN
			GVL_TWO_PALLET.auiCommand[uiTwin] := 16;
		END_IF;
	END_IF;

	// Единственное место преобразования транспортных номеров HMI в интерфейс FB.
	astTwinCommand[uiTwin].xEnable := GVL_TWO_PALLET.auiCommand[uiTwin] = UINT#1;
	astTwinCommand[uiTwin].xConfirm := GVL_TWO_PALLET.auiCommand[uiTwin] = UINT#2;
	astTwinCommand[uiTwin].xStart := GVL_TWO_PALLET.auiCommand[uiTwin] = UINT#27;
	astTwinCommand[uiTwin].xRejectStart := GVL_TWO_PALLET.auiCommand[uiTwin] = UINT#28;
	astTwinCommand[uiTwin].xDisable := GVL_TWO_PALLET.auiCommand[uiTwin] = UINT#3;
	astTwinCommand[uiTwin].xSwap := GVL_TWO_PALLET.auiCommand[uiTwin] = UINT#4;
	astTwinCommand[uiTwin].xPowerOn := GVL_TWO_PALLET.auiCommand[uiTwin] = UINT#5;
	astTwinCommand[uiTwin].xPowerOff := GVL_TWO_PALLET.auiCommand[uiTwin] = UINT#6;
	astTwinCommand[uiTwin].xDriveReset := GVL_TWO_PALLET.auiCommand[uiTwin] = UINT#7;
	astTwinCommand[uiTwin].xHome := GVL_TWO_PALLET.auiCommand[uiTwin] = UINT#8;
	astTwinCommand[uiTwin].xLower := GVL_TWO_PALLET.auiCommand[uiTwin] = UINT#9;
	astTwinCommand[uiTwin].xRaise := GVL_TWO_PALLET.auiCommand[uiTwin] = UINT#10;
	astTwinCommand[uiTwin].xSelectPallet := (GVL_TWO_PALLET.auiCommand[uiTwin] = UINT#11)
		OR (GVL_TWO_PALLET.auiCommand[uiTwin] = UINT#12);
	astTwinCommand[uiTwin].xLockIn := GVL_TWO_PALLET.auiCommand[uiTwin] = UINT#29;
	astTwinCommand[uiTwin].xLockOut := GVL_TWO_PALLET.auiCommand[uiTwin] = UINT#30;
	astTwinCommand[uiTwin].xStopIn := GVL_TWO_PALLET.auiCommand[uiTwin] = UINT#31;
	astTwinCommand[uiTwin].xStopOut := GVL_TWO_PALLET.auiCommand[uiTwin] = UINT#32;
	astTwinCommand[uiTwin].xMoveToExchange := GVL_TWO_PALLET.auiCommand[uiTwin] = UINT#13;
	astTwinCommand[uiTwin].xMoveToWork := GVL_TWO_PALLET.auiCommand[uiTwin] = UINT#14;
	astTwinCommand[uiTwin].xStop := GVL_TWO_PALLET.auiCommand[uiTwin] = UINT#15;
	astTwinCommand[uiTwin].xReset := GVL_TWO_PALLET.auiCommand[uiTwin] = UINT#16;
	astTwinCommand[uiTwin].xJogPositive := GVL_TWO_PALLET.auiCommand[uiTwin] = UINT#17;
	astTwinCommand[uiTwin].xJogNegative := GVL_TWO_PALLET.auiCommand[uiTwin] = UINT#18;
	astTwinCommand[uiTwin].xJogRelease := GVL_TWO_PALLET.auiCommand[uiTwin] = UINT#19;
	astTwinCommand[uiTwin].xTeachOperator := GVL_TWO_PALLET.auiCommand[uiTwin] = UINT#25;
	astTwinCommand[uiTwin].xTeachWork := GVL_TWO_PALLET.auiCommand[uiTwin] = UINT#26;
	astTwinCommand[uiTwin].uiPallet := GVL_TWO_PALLET.auiValue[uiTwin];
	IF GVL_TWO_PALLET.auiCommand[uiTwin] = UINT#11 THEN
		astTwinCommand[uiTwin].uiPallet := UINT#1;
	ELSIF GVL_TWO_PALLET.auiCommand[uiTwin] = UINT#12 THEN
		astTwinCommand[uiTwin].uiPallet := UINT#2;
	END_IF;
	astTwinCommand[uiTwin].udiRevision := GVL_TWO_PALLET.audiRevision[uiTwin];

	IF xTestInitializePulse AND (GVL_CELL_SETTINGS.eTestEnvironment = E_CELL_TEST_ENVIRONMENT.SIMULATION) THEN
		astTwinCommand[uiTwin].xEnable := GVL_HMI.stTestScenario.axMagazineEnabled[uiTwin];
		astTwinCommand[uiTwin].xDisable := NOT GVL_HMI.stTestScenario.axMagazineEnabled[uiTwin];
	END_IF;

	// Фактическая операция включает удерживаемый запрос и завершение Disable.
	// Предпочтение возврата удерживает только автообмен до последнего PUT.
	// Повторное включение и ручная наладка зависят от фактической операции.
	// Занятость другого магазина/станка сама по себе не запрещает правку инвентаря.
	xTwinRobotOperation := GVL_MAGAZINE.astPartStatus[uiTwin].xBusy
		OR GVL_MAGAZINE.astPartStatus[uiTwin].xDisablePending
		OR GVL_MAGAZINE.astAutoCommand[uiTwin].xExecute
		OR GVL_MAGAZINE.astCommand[uiTwin].xExecute
		OR ((GVL_ROBOT.Status.xBusy OR xMotionBusy)
			AND (GVL_ROBOT.Status.uiMagazineContext = uiTwin))
		OR ((GVL_CELL_MANAGER.Status.uiActiveMagazine = uiTwin)
			AND ((GVL_CELL_MANAGER.Diag.eState = E_CELL_STATE.MAGAZINE)
				OR (GVL_CELL_MANAGER.Diag.eState = E_CELL_STATE.RELEASE_MAGAZINE)));
	// Для обмена важна занятость только этого магазина. Точка и состояние
	// интерфейса робота после инициализации могут быть неизвестны.
	xTwinRobotSwapWindow := NOT xTwinRobotOperation
		AND (CELL_MANAGER.uiReturnMagazine <> uiTwin);
	xTwinOtherLoaded := FALSE;
	xTwinRobotHasBlank := TRUE; // Неизвестная роль палеты запрещает автоматический обмен
	xTwinOtherHasBlank := FALSE;
	xTwinInventoryEditPending := xTwinInventoryCommand
		AND (stTwinRequest.uiMagazine = uiTwin)
		AND (stTwinRequest.uiCommand >= UINT#21)
		AND (stTwinRequest.uiCommand <= UINT#24);
	IF (GVL_TWO_PALLET.astStatus[uiTwin].uiRobotPallet >= UINT#1)
		AND (GVL_TWO_PALLET.astStatus[uiTwin].uiRobotPallet <= UINT#2) THEN
		uiTwinPallet := UINT#3 - GVL_TWO_PALLET.astStatus[uiTwin].uiRobotPallet;
		xTwinOtherLoaded := GVL_TWO_PALLET.astStore[uiTwin].axLoaded[uiTwinPallet];
		xTwinRobotHasBlank := FALSE;
		FOR uiTwinSlot := UINT#1 TO UINT#96 DO
			IF GVL_TWO_PALLET.astStore[uiTwin].astPallet[GVL_TWO_PALLET.astStatus[uiTwin].uiRobotPallet].aSlots[uiTwinSlot].xInPosition
			AND (GVL_TWO_PALLET.astStore[uiTwin].astPallet[GVL_TWO_PALLET.astStatus[uiTwin].uiRobotPallet].aSlots[uiTwinSlot].eDetailType = E_DETAIL_TYPE.BLANK) THEN
				xTwinRobotHasBlank := TRUE;
			END_IF;
			IF GVL_TWO_PALLET.astStore[uiTwin].astPallet[uiTwinPallet].aSlots[uiTwinSlot].xInPosition
			AND (GVL_TWO_PALLET.astStore[uiTwin].astPallet[uiTwinPallet].aSlots[uiTwinSlot].eDetailType = E_DETAIL_TYPE.BLANK) THEN
				xTwinOtherHasBlank := TRUE;
			END_IF;
		END_FOR;
	END_IF;
	// Finished сохраняет ожидание оператора. Ранний запрос отменяемый: при утрате
	// подготовки палета остаётся доступной для выгрузки, её Finished не защёлкивается.
	// Сканируем фактические карты, включая заготовки неподходящих сейчас типов.
	axTwinAutoSwapPending[uiTwin] := (GVL_TWO_PALLET.uiMode = UINT#1)
		AND GVL_CELL_MANAGER.Status.xRunning
		AND NOT GVL_CELL_MANAGER.Status.xStopPending
		AND NOT GVL_CELL_CONTROL.xStop
		AND NOT GVL_CELL_CONTROL.xManual
		AND NOT xTwinRobotHasBlank
		AND (GVL_MAGAZINE.astPartStatus[uiTwin].xFinished
			OR (xTwinAutoSwapEnabled AND xTwinOtherLoaded AND xTwinOtherHasBlank
				AND NOT xTwinInventoryEditPending AND xTwinRobotSwapWindow))
		AND NOT astTwinCommand[uiTwin].xDisable
		AND NOT astTwinCommand[uiTwin].xStop;
	uiTwinRobotPalletBefore := GVL_TWO_PALLET.astStatus[uiTwin].uiRobotPallet;
	TWIN[uiTwin](
		xSelected := GVL_TWO_PALLET.uiMode = 1,
		xManual := GVL_CELL_CONTROL.xManual AND NOT GVL_CELL_MANAGER.Status.xRunning,
		xSafe := CELL_SAFETY.Status.xReady AND NOT GVL_CELL_CONTROL.xGlobalError AND NOT GVL_HMI.xIoEmergencyStopActive
			AND CELL_SAFETY.astEnclosureDoorStatus[uiTwin * 2 - 1].xLocked
			AND CELL_SAFETY.astEnclosureDoorStatus[uiTwin * 2].xLocked
			AND NOT CELL_SAFETY.astEnclosureDoorStatus[uiTwin * 2 - 1].xUnlockOutput
			AND NOT CELL_SAFETY.astEnclosureDoorStatus[uiTwin * 2].xUnlockOutput,
		xRobotSwapWindow := xTwinRobotSwapWindow,
		xRobotOperation := xTwinRobotOperation,
		xPointsConfigured := axMagazinePointsReady[uiTwin],
		xRobotGeometryReady := NOT GVL_HMI.xModbusMode AND axMagazinePointsReady[uiTwin],
		xRobotMagazineReady := GVL_MAGAZINE.astPartStatus[uiTwin].xEnableCheckNoError
			AND GVL_MAGAZINE.astPartStatus[uiTwin].xEnableCheckGeometry,
		xConnection := xHmiConnectionAlive,
		xStopRequest := GVL_CELL_CONTROL.xStop OR xIoManualActive OR GVL_HMI.astMagazineCommand[uiTwin].xStop OR GVL_TWO_PALLET.xModeChanged,
		xAutoSwap := axTwinAutoSwapPending[uiTwin] AND xTwinAutoSwapEnabled
			AND xTwinOtherLoaded AND xTwinOtherHasBlank AND NOT xTwinInventoryEditPending,
		xOtherLoaded := xTwinOtherLoaded,
		xActivePalletEditAllowed := NOT xTwinRobotOperation,
		xConfigurationChanged := axTwinConfigurationChanged[uiTwin],
        xIoPneumaticOverride := axIoMagazineInvalidated[uiTwin],
		xExternalCommandRejected := axTwinExternalCommandRejected[uiTwin],
		Command := astTwinCommand[uiTwin],
		Config := GVL_TWO_PALLET.astActiveConfig[uiTwin], Input := GVL_TWO_PALLET.astInput[uiTwin],
		Status => GVL_TWO_PALLET.astStatus[uiTwin],
		Diag => GVL_TWO_PALLET.astDiag[uiTwin],
		Error => GVL_TWO_PALLET.astError[uiTwin],
		Output => GVL_TWO_PALLET.astOutput[uiTwin]);
    axIoMagazineInvalidated[uiTwin] := FALSE;
	// Блокировка относится только к этому магазину и удерживается до полного
	// окончания механического обмена, включая последний скан Completed.
	axTwinMagazineExchangeInProgress[uiTwin] := GVL_TWO_PALLET.astStatus[uiTwin].xBusy
		OR GVL_TWO_PALLET.astStatus[uiTwin].xCompleted;
	GVL_TWO_PALLET.astStatus[uiTwin].xAutoSwapEnabled := xTwinAutoSwapEnabled;
	// После Stop/Disable или аварии ожидание обмена не удерживает планировщик.
	axTwinAutoSwapPending[uiTwin] := axTwinAutoSwapPending[uiTwin]
		AND NOT GVL_TWO_PALLET.astStatus[uiTwin].xError;
	axTwinConfigurationChanged[uiTwin] := FALSE;
	axTwinExternalCommandRejected[uiTwin] := FALSE;
	IF GVL_TWO_PALLET.astOutput[uiTwin].xTeachOperator THEN
		IF GVL_CELL_SETTINGS.eTestEnvironment = E_CELL_TEST_ENVIRONMENT.SIMULATION THEN
			GVL_TWO_PALLET.astSimulationConfig[uiTwin].lrExchange := GVL_TWO_PALLET.astInput[uiTwin].lrPosition;
		ELSE
			GVL_TWO_PALLET.astConfig[uiTwin].lrExchange := GVL_TWO_PALLET.astInput[uiTwin].lrPosition;
		END_IF;
		axTwinConfigurationChanged[uiTwin] := TRUE;
	END_IF;
	IF GVL_TWO_PALLET.astOutput[uiTwin].xTeachWork THEN
		IF GVL_TWO_PALLET.astStatus[uiTwin].uiSelected = UINT#1 THEN
			IF GVL_CELL_SETTINGS.eTestEnvironment = E_CELL_TEST_ENVIRONMENT.SIMULATION THEN
				GVL_TWO_PALLET.astSimulationConfig[uiTwin].lrWorkP1 := GVL_TWO_PALLET.astInput[uiTwin].lrPosition;
			ELSE
				GVL_TWO_PALLET.astConfig[uiTwin].lrWorkP1 := GVL_TWO_PALLET.astInput[uiTwin].lrPosition;
			END_IF;
		ELSIF GVL_TWO_PALLET.astStatus[uiTwin].uiSelected = UINT#2 THEN
			IF GVL_CELL_SETTINGS.eTestEnvironment = E_CELL_TEST_ENVIRONMENT.SIMULATION THEN
				GVL_TWO_PALLET.astSimulationConfig[uiTwin].lrWorkP2 := GVL_TWO_PALLET.astInput[uiTwin].lrPosition;
			ELSE
				GVL_TWO_PALLET.astConfig[uiTwin].lrWorkP2 := GVL_TWO_PALLET.astInput[uiTwin].lrPosition;
			END_IF;
		END_IF;
		axTwinConfigurationChanged[uiTwin] := TRUE;
	END_IF;
	// RunCellControl ниже должен видеть запрет уже в скане начала обмена.
	IF GVL_TWO_PALLET.uiMode = 1 THEN
		GVL_MAGAZINE.astStatus[uiTwin].xReady := GVL_MAGAZINE.astPartStatus[uiTwin].xReady
			AND GVL_TWO_PALLET.astStatus[uiTwin].xReady;
		GVL_MAGAZINE.astStatus[uiTwin].xBusy := GVL_MAGAZINE.astPartStatus[uiTwin].xBusy
			OR GVL_TWO_PALLET.astStatus[uiTwin].xBusy;
		GVL_MAGAZINE.astStatus[uiTwin].xEnabled := GVL_TWO_PALLET.astStatus[uiTwin].xEnabled;
	END_IF;
	IF GVL_TWO_PALLET.astStatus[uiTwin].xCompleted THEN
		GVL_TWO_PALLET.astStore[uiTwin].axLoaded[1] := FALSE;
		GVL_TWO_PALLET.astStore[uiTwin].axLoaded[2] := FALSE;
		axTwinStoreChanged[uiTwin] := TRUE;
		axMagazineInventoryChanged[uiTwin] := TRUE;
	END_IF;
	// Ручное восстановление может сменить учётную роль без команды обмена.
	IF uiTwinRobotPalletBefore <> GVL_TWO_PALLET.astStatus[uiTwin].uiRobotPallet THEN
		GVL_TWO_PALLET.astStore[uiTwin].axLoaded[1] := FALSE;
		GVL_TWO_PALLET.astStore[uiTwin].axLoaded[2] := FALSE;
		axTwinStoreChanged[uiTwin] := TRUE;
		axMagazineInventoryChanged[uiTwin] := TRUE;
	END_IF;
	// Ручная смена расходует прежнее подтверждение уже при принятии команды.
	IF astTwinCommand[uiTwin].xSwap AND GVL_TWO_PALLET.astStatus[uiTwin].xCommandAccepted THEN
		GVL_TWO_PALLET.astStore[uiTwin].axLoaded[1] := FALSE;
		GVL_TWO_PALLET.astStore[uiTwin].axLoaded[2] := FALSE;
		axTwinStoreChanged[uiTwin] := TRUE;
	END_IF;
	IF (uiTwinRequestResult = 2) AND (stTwinRequest.uiMagazine = uiTwin)
		AND (((stTwinRequest.uiCommand >= 1) AND (stTwinRequest.uiCommand <= 19))
			OR ((stTwinRequest.uiCommand >= 25) AND (stTwinRequest.uiCommand <= 32)))
		AND GVL_TWO_PALLET.astStatus[uiTwin].xCommandAccepted THEN uiTwinRequestResult := 1; END_IF;
END_FOR;

IF xTwinInventoryCommand THEN
	uiTwin := stTwinRequest.uiMagazine;
	uiTwinPallet := stTwinRequest.uiValue;
	IF stTwinRequest.uiCommand = UINT#24 THEN
		IF GVL_TWO_PALLET.astStatus[uiTwin].xConfigAllowed
			AND stTwinRequest.Config.xSignalPatternsConfigured
			AND TWIN[uiTwin].IsSignalConfigurationValid(
				uiP1Signals := stTwinRequest.Config.uiP1Signals,
				uiP2Signals := stTwinRequest.Config.uiP2Signals) THEN
			IF GVL_CELL_SETTINGS.eTestEnvironment = E_CELL_TEST_ENVIRONMENT.SIMULATION THEN
				GVL_TWO_PALLET.astSimulationConfig[uiTwin] := stTwinRequest.Config;
			ELSE
				GVL_TWO_PALLET.astConfig[uiTwin] := stTwinRequest.Config;
			END_IF;
			axTwinConfigurationChanged[uiTwin] := TRUE;
			uiTwinRequestResult := UINT#1;
		END_IF;
	ELSIF ((uiTwinPallet = 1) AND GVL_TWO_PALLET.astStatus[uiTwin].xEdit1Allowed)
		OR ((uiTwinPallet = 2) AND GVL_TWO_PALLET.astStatus[uiTwin].xEdit2Allowed) THEN
		CASE stTwinRequest.uiCommand OF
			20:
				IF GVL_TWO_PALLET.astStatus[uiTwin].xLoadAllowed
					AND (uiTwinPallet <> GVL_TWO_PALLET.astStatus[uiTwin].uiRobotPallet) THEN
					axTwinStoreChanged[uiTwin] := TRUE;
					GVL_TWO_PALLET.astStore[uiTwin].axLoaded[uiTwinPallet] := TRUE;
					uiTwinRequestResult := 1;
				END_IF;
			21, 22:
				FOR uiTwinSlot := 1 TO 96 DO
					GVL_TWO_PALLET.astStore[uiTwin].astPallet[uiTwinPallet].aSlots[uiTwinSlot].xInPosition := stTwinRequest.uiCommand = 22;
					GVL_TWO_PALLET.astStore[uiTwin].astPallet[uiTwinPallet].aSlots[uiTwinSlot].eDetailType := E_DETAIL_TYPE.NONE;
					GVL_TWO_PALLET.astStore[uiTwin].astPallet[uiTwinPallet].aSlots[uiTwinSlot].uiProductType := 0;
					IF stTwinRequest.uiCommand = 22 THEN
						GVL_TWO_PALLET.astStore[uiTwin].astPallet[uiTwinPallet].aSlots[uiTwinSlot].eDetailType := E_DETAIL_TYPE.BLANK;
						GVL_TWO_PALLET.astStore[uiTwin].astPallet[uiTwinPallet].aSlots[uiTwinSlot].uiProductType := GVL_MULTI_TYPE.Config.auiSlotType[uiTwinSlot];
					END_IF;
				END_FOR;
				axTwinStoreChanged[uiTwin] := TRUE;
				GVL_TWO_PALLET.astStore[uiTwin].axLoaded[uiTwinPallet] := FALSE; uiTwinRequestResult := 1;
			23:
				IF (stTwinRequest.uiSlot >= 1) AND (stTwinRequest.uiSlot <= 96) AND (stTwinRequest.uiContent <= 2)
					AND ((stTwinRequest.uiContent = 0) OR ((stTwinRequest.uiProductType >= 1) AND (stTwinRequest.uiProductType <= GVL_MULTI_TYPE.Config.uiTypeCount))) THEN
					uiTwinSlot := stTwinRequest.uiSlot;
					GVL_TWO_PALLET.astStore[uiTwin].astPallet[uiTwinPallet].aSlots[uiTwinSlot].xInPosition := stTwinRequest.uiContent <> 0;
					CASE stTwinRequest.uiContent OF
						0: GVL_TWO_PALLET.astStore[uiTwin].astPallet[uiTwinPallet].aSlots[uiTwinSlot].eDetailType := E_DETAIL_TYPE.NONE;
						1: GVL_TWO_PALLET.astStore[uiTwin].astPallet[uiTwinPallet].aSlots[uiTwinSlot].eDetailType := E_DETAIL_TYPE.BLANK;
						2: GVL_TWO_PALLET.astStore[uiTwin].astPallet[uiTwinPallet].aSlots[uiTwinSlot].eDetailType := E_DETAIL_TYPE.DETAIL;
					END_CASE;
					GVL_TWO_PALLET.astStore[uiTwin].astPallet[uiTwinPallet].aSlots[uiTwinSlot].uiProductType := stTwinRequest.uiProductType;
					axTwinStoreChanged[uiTwin] := TRUE;
					GVL_TWO_PALLET.astStore[uiTwin].axLoaded[uiTwinPallet] := FALSE; uiTwinRequestResult := 1;
				END_IF;
		END_CASE;
		// Загрузка/редактирование палеты у оператора не отменяет завершение рабочей.
		IF (uiTwinRequestResult = UINT#1)
			AND (stTwinRequest.uiCommand >= UINT#21)
			AND (stTwinRequest.uiCommand <= UINT#23)
			AND (uiTwinPallet = GVL_TWO_PALLET.astStatus[uiTwin].uiRobotPallet) THEN
			axMagazineInventoryChanged[uiTwin] := TRUE;
		END_IF;
	END_IF;
END_IF;
IF uiTwinRequestResult <> 0 THEN
	GVL_HMI.uiTwinResult := uiTwinRequestResult;
	GVL_HMI.udiTwinAckSeq := udiTwinSnapshot;
	IF uiTwinRequestResult <> 1 THEN
		uiTwin := LIMIT(UINT#1, stTwinRequest.uiMagazine, UINT#2);
		// Команды механизма 1..19 и 25..28 уже формируют предупреждение внутри FB в этом же скане.
		IF GVL_TWO_PALLET.auiCommand[uiTwin] <> stTwinRequest.uiCommand THEN
			axTwinExternalCommandRejected[uiTwin] := TRUE;
		END_IF;
	END_IF;
END_IF;

GVL_CELL_SETTINGS.MagazineRows := 12;
GVL_CELL_SETTINGS.MagazineColumns := 10;
IF GVL_TWO_PALLET.uiMode = 1 THEN GVL_CELL_SETTINGS.MagazineRows := 12; GVL_CELL_SETTINGS.MagazineColumns := 8; END_IF;
GVL_HMI.MagazineRows := GVL_CELL_SETTINGS.MagazineRows;
GVL_HMI.MagazineColumns := GVL_CELL_SETTINGS.MagazineColumns;
FOR uiTwin := 1 TO 2 DO
	IF GVL_TWO_PALLET.uiMode = 1 THEN
		uiTwinPallet := GVL_TWO_PALLET.astStatus[uiTwin].uiRobotPallet;
		IF (uiTwinPallet < UINT#1) OR (uiTwinPallet > UINT#2) THEN
			uiTwinPallet := UINT#1;
		END_IF;
        IF axMagazineInventoryChanged[uiTwin] THEN
            GVL_DETAIL.astMagazine[uiTwin] := GVL_TWO_PALLET.astStore[uiTwin].astPallet[uiTwinPallet];
        END_IF;
	END_IF;
END_FOR;

(* ---- PLC_PRG.RunTwoPalletAxis.st ---- *)
METHOD PRIVATE RunTwoPalletAxis

// --- BEGIN IMPLEMENTATION ---

// Magazine_1/2 — точки привязки Motion: в NORMAL настроить реальные оси EtherCAT.
// MC_Home запускает поиск дома в серводрайвере; FB_AXIS ждёт его Done.
// Ссылки назначаются каждый скан до проверки __ISVALIDREF и вызова FB_AXIS.
GVL_TWO_PALLET.Axis1 REF= Magazine_1;
GVL_TWO_PALLET.Axis2 REF= Magazine_2;
GVL_TWO_PALLET.astInput[1].xAxisBound := __ISVALIDREF(GVL_TWO_PALLET.Axis1);
GVL_TWO_PALLET.astInput[2].xAxisBound := __ISVALIDREF(GVL_TWO_PALLET.Axis2);
FOR uiTwin := 1 TO 2 DO
	GVL_TWO_PALLET.astAxis[uiTwin].Command.xEnable := GVL_TWO_PALLET.astOutput[uiTwin].xPowerOn;
	GVL_TWO_PALLET.astAxis[uiTwin].Command.xDisable := GVL_TWO_PALLET.astOutput[uiTwin].xPowerOff
		OR (GVL_TWO_PALLET.uiMode = 0);
	GVL_TWO_PALLET.astAxis[uiTwin].Command.xPowerPermit := (GVL_TWO_PALLET.uiMode = 1)
		AND CELL_SAFETY.Status.xReady AND GVL_TWO_PALLET.astInput[uiTwin].xIoMapped;
	GVL_TWO_PALLET.astAxis[uiTwin].Command.xGlobalError := GVL_CELL_CONTROL.xGlobalError;
	GVL_TWO_PALLET.astAxis[uiTwin].Command.xResetAllError := GVL_TWO_PALLET.astOutput[uiTwin].xDriveReset;
	GVL_TWO_PALLET.astAxis[uiTwin].Command.xStop := GVL_TWO_PALLET.astOutput[uiTwin].xStop OR GVL_HMI.xIoEmergencyStopActive;
	GVL_TWO_PALLET.astAxis[uiTwin].Command.xHome := GVL_TWO_PALLET.astOutput[uiTwin].xHome;
	GVL_TWO_PALLET.astAxis[uiTwin].Command.xMoveAbsolute := GVL_TWO_PALLET.astOutput[uiTwin].xMove;
	GVL_TWO_PALLET.astAxis[uiTwin].Command.xJogPositive := GVL_TWO_PALLET.astOutput[uiTwin].xJogPositive;
	GVL_TWO_PALLET.astAxis[uiTwin].Command.xJogNegative := GVL_TWO_PALLET.astOutput[uiTwin].xJogNegative;
	GVL_TWO_PALLET.astAxis[uiTwin].MotionParam.lrTargetPosition := GVL_TWO_PALLET.astOutput[uiTwin].lrTarget;
	GVL_TWO_PALLET.astAxis[uiTwin].MotionParam.lrHomePosition := GVL_TWO_PALLET.astActiveConfig[uiTwin].lrHome;
	GVL_TWO_PALLET.astAxis[uiTwin].MotionParam.lrVelocity := GVL_TWO_PALLET.astActiveConfig[uiTwin].lrVelocity;
	GVL_TWO_PALLET.astAxis[uiTwin].MotionParam.lrAcceleration := GVL_TWO_PALLET.astActiveConfig[uiTwin].lrAcceleration;
	GVL_TWO_PALLET.astAxis[uiTwin].MotionParam.lrDeceleration := GVL_TWO_PALLET.astActiveConfig[uiTwin].lrDeceleration;
	GVL_TWO_PALLET.astAxis[uiTwin].MotionParam.lrJerk := GVL_TWO_PALLET.astActiveConfig[uiTwin].lrJerk;
	GVL_TWO_PALLET.astAxis[uiTwin].Timeouts := GVL_CELL_SETTINGS.stAxisTimeouts;
	GVL_TWO_PALLET.astAxis[uiTwin].Timeouts.tHomeTimeout := GVL_TWO_PALLET.astActiveConfig[uiTwin].tHome;
	GVL_TWO_PALLET.astAxis[uiTwin].Timeouts.tMoveTimeout := GVL_TWO_PALLET.astActiveConfig[uiTwin].tMove;
END_FOR;
IF __ISVALIDREF(GVL_TWO_PALLET.Axis1) THEN
	TWIN_AXIS_1(Axis := GVL_TWO_PALLET.Axis1, AxisData := GVL_TWO_PALLET.astAxis[1],
		xResetPermit := GVL_CELL_CONTROL.xManual AND NOT GVL_CELL_MANAGER.Status.xRunning);
END_IF;
IF __ISVALIDREF(GVL_TWO_PALLET.Axis2) THEN
	TWIN_AXIS_2(Axis := GVL_TWO_PALLET.Axis2, AxisData := GVL_TWO_PALLET.astAxis[2],
		xResetPermit := GVL_CELL_CONTROL.xManual AND NOT GVL_CELL_MANAGER.Status.xRunning);
END_IF;
FOR uiTwin := 1 TO 2 DO
	GVL_TWO_PALLET.astInput[uiTwin].xPowered := GVL_TWO_PALLET.astAxis[uiTwin].Status.xPowered;
	GVL_TWO_PALLET.astInput[uiTwin].xHomed := GVL_TWO_PALLET.astAxis[uiTwin].Status.xHomed;
	GVL_TWO_PALLET.astInput[uiTwin].xStandstill := GVL_TWO_PALLET.astAxis[uiTwin].Status.xStandstill;
	GVL_TWO_PALLET.astInput[uiTwin].xDriveError := GVL_TWO_PALLET.astAxis[uiTwin].Status.xError;
	GVL_TWO_PALLET.astInput[uiTwin].xMotionDone := GVL_TWO_PALLET.astAxis[uiTwin].Status.xDone;
	GVL_TWO_PALLET.astInput[uiTwin].lrPosition := GVL_TWO_PALLET.astAxis[uiTwin].Status.lrActualPosition;
	TWIN_SIM[uiTwin](
		xEnable := (GVL_TWO_PALLET.uiMode = UINT#1)
			AND (GVL_CELL_SETTINGS.eTestEnvironment = E_CELL_TEST_ENVIRONMENT.SIMULATION),
		uiP1Signals := GVL_TWO_PALLET.astActiveConfig[uiTwin].uiP1Signals,
		Command := GVL_TWO_PALLET.astOutput[uiTwin]);
	IF (GVL_TWO_PALLET.uiMode = UINT#1)
		AND (GVL_CELL_SETTINGS.eTestEnvironment = E_CELL_TEST_ENVIRONMENT.SIMULATION) THEN
		GVL_TWO_PALLET.astInput[uiTwin].xIoMapped := TRUE;
		GVL_TWO_PALLET.astInput[uiTwin].xLiftDown := TWIN_SIM[uiTwin].xLiftDown;
		GVL_TWO_PALLET.astInput[uiTwin].xLiftUp := TWIN_SIM[uiTwin].xLiftUp;
		GVL_TWO_PALLET.astInput[uiTwin].xLockIn := TWIN_SIM[uiTwin].xLockIn;
		GVL_TWO_PALLET.astInput[uiTwin].xLockOut := TWIN_SIM[uiTwin].xLockOut;
		GVL_TWO_PALLET.astInput[uiTwin].xStopIn := TWIN_SIM[uiTwin].xStopIn;
		GVL_TWO_PALLET.astInput[uiTwin].xStopOut := TWIN_SIM[uiTwin].xStopOut;
		GVL_TWO_PALLET.astInput[uiTwin].xLimitNegative := FALSE;
		GVL_TWO_PALLET.astInput[uiTwin].xLimitPositive := FALSE;
		GVL_TWO_PALLET.astInput[uiTwin].xHomeSensor := GVL_TWO_PALLET.astInput[uiTwin].xHomed
			AND (ABS(GVL_TWO_PALLET.astInput[uiTwin].lrPosition
				- GVL_TWO_PALLET.astActiveConfig[uiTwin].lrHome)
				<= GVL_TWO_PALLET.astActiveConfig[uiTwin].lrTolerance);
		axTwinSimIoOwned[uiTwin] := TRUE;
	ELSIF axTwinSimIoOwned[uiTwin]
	AND (GVL_CELL_SETTINGS.eTestEnvironment <> E_CELL_TEST_ENVIRONMENT.NORMAL) THEN
		// После выхода из виртуальной среды не оставляем её герконы как реальные.
		GVL_TWO_PALLET.astInput[uiTwin].xIoMapped := FALSE;
		GVL_TWO_PALLET.astInput[uiTwin].xLiftDown := FALSE;
		GVL_TWO_PALLET.astInput[uiTwin].xLiftUp := FALSE;
		GVL_TWO_PALLET.astInput[uiTwin].xLockIn := FALSE;
		GVL_TWO_PALLET.astInput[uiTwin].xLockOut := FALSE;
		GVL_TWO_PALLET.astInput[uiTwin].xStopIn := FALSE;
		GVL_TWO_PALLET.astInput[uiTwin].xStopOut := FALSE;
		GVL_TWO_PALLET.astInput[uiTwin].xLimitNegative := FALSE;
		GVL_TWO_PALLET.astInput[uiTwin].xLimitPositive := FALSE;
		GVL_TWO_PALLET.astInput[uiTwin].xHomeSensor := FALSE;
		axTwinSimIoOwned[uiTwin] := FALSE;
	END_IF;
	IF GVL_CELL_SETTINGS.eTestEnvironment = E_CELL_TEST_ENVIRONMENT.NORMAL THEN
		// ReadPhysicalInputs уже заменил виртуальные герконы в начале скана.
		// Концевики и датчик дома заведены в драйвер, не в DI ячейки. Эти legacy-
		// поля не имитируют PDO; результат Home приходит выше через xHomed/xMotionDone.
		GVL_TWO_PALLET.astInput[uiTwin].xLimitNegative := FALSE;
		GVL_TWO_PALLET.astInput[uiTwin].xLimitPositive := FALSE;
		GVL_TWO_PALLET.astInput[uiTwin].xHomeSensor := FALSE;
		axTwinSimIoOwned[uiTwin] := FALSE;
	END_IF;
END_FOR;

(* ---- PLC_PRG.SetApplicationDefaults.st ---- *)
METHOD PRIVATE SetApplicationDefaults

// --- BEGIN IMPLEMENTATION ---

// При старте PLC ячейка всегда включается в ручном режиме: автоматический цикл
// требует явного переключения оператором. Однократный флаг также повторно
// применяет безопасные значения при Online Change, когда initializer GVL
// может не перезаписать уже существующее значение. Инициализация выполняется до
// RunCellControl, чтобы автомат не увидел прежние настройки даже на один цикл.
IF NOT xApplicationStartupInitialized THEN
	GVL_CELL_CONTROL.xManual := TRUE;
	FOR uiMachine := 1 TO 3 DO
		GVL_HMI.axMachineUsed[uiMachine] := FALSE;
	END_FOR;
	// RETAIN uiMode переживает перезапуск PLC, поэтому явно выбираем двухпалетный
	// тип на старте. При реальной смене типа старые базы магазинов недействительны.
	IF GVL_TWO_PALLET.uiMode <> UINT#1 THEN
		GVL_TWO_PALLET.uiMode := UINT#1;
		InvalidateMagazineCalibration(uiMagazine := UINT#1);
		InvalidateMagazineCalibration(uiMagazine := UINT#2);
		xPointTableReady := FALSE;
	END_IF;
	GVL_CELL_SETTINGS.eTestEnvironment := E_CELL_TEST_ENVIRONMENT.SIMULATION;
	xApplicationStartupInitialized := TRUE;
END_IF;

// При первом запуске этой схемы намеренно отбрасываем прежние инженерные
// координаты. Нулевая скорость и xConfigured=FALSE не позволяют принять
// нулевую точку за пригодную для движения.
IF Persistent_Value.udiPointStorageVersion <> GVL_POINT.udiExpectedPointStorageVersion THEN
	FOR uiPointEditorIndex := UINT#1 TO INT_TO_UINT(GVL_POINT.iPersistentPointCapacity) DO
		Persistent_Value.astRetainPoints[uiPointEditorIndex].Name := '';
		Persistent_Value.astRetainPoints[uiPointEditorIndex].X := 0.0;
		Persistent_Value.astRetainPoints[uiPointEditorIndex].Y := 0.0;
		Persistent_Value.astRetainPoints[uiPointEditorIndex].Z := 0.0;
		Persistent_Value.astRetainPoints[uiPointEditorIndex].MagazineSafeZ := 0.0;
		Persistent_Value.astRetainPoints[uiPointEditorIndex].MagazineChangeZ := 0.0;
		Persistent_Value.astRetainPoints[uiPointEditorIndex].SpeedFactor := 0.0;
		Persistent_Value.astRetainPoints[uiPointEditorIndex].xConfigured := FALSE;
	END_FOR;
	Persistent_Value.udiPointStorageVersion := GVL_POINT.udiExpectedPointStorageVersion;
END_IF;

// Единственное соответствие компактного редакторского индекса, стабильного
// E_POINT_NAME и прежнего индекса Persistent-массива. Три legacy-точки INSIDE
// пропущены; рецепты станков их не используют.
xPointTableReady := TRUE;
// Базы ГК хранятся у владельца GVL_GEOMETRY_CONTROL, отдельно от прежних 15
// Persistent-позиций. Их добавление не сбрасывает уже сохранённые точки.
FOR uiPointEditorIndex := UINT#1 TO INT_TO_UINT(GVL_POINT.iRequiredPointCount) DO
	uiPointStorageIndex := UINT#0;
	CASE uiPointEditorIndex OF
		UINT#1: ePointEditorName := E_POINT_NAME.MACHINE_1_ABOVE; uiPointStorageIndex := UINT#1;
		UINT#2: ePointEditorName := E_POINT_NAME.MACHINE_1_CHUCK_APROACH; uiPointStorageIndex := UINT#3;
		UINT#3: ePointEditorName := E_POINT_NAME.MACHINE_1_CHUCK_POSITION; uiPointStorageIndex := UINT#4;
		UINT#4: ePointEditorName := E_POINT_NAME.MACHINE_2_ABOVE; uiPointStorageIndex := UINT#5;
		UINT#5: ePointEditorName := E_POINT_NAME.MACHINE_2_CHUCK_APROACH; uiPointStorageIndex := UINT#7;
		UINT#6: ePointEditorName := E_POINT_NAME.MACHINE_2_CHUCK_POSITION; uiPointStorageIndex := UINT#8;
		UINT#7: ePointEditorName := E_POINT_NAME.MACHINE_3_ABOVE; uiPointStorageIndex := UINT#9;
		UINT#8: ePointEditorName := E_POINT_NAME.MACHINE_3_CHUCK_APROACH; uiPointStorageIndex := UINT#11;
		UINT#9: ePointEditorName := E_POINT_NAME.MACHINE_3_CHUCK_POSITION; uiPointStorageIndex := UINT#12;
		UINT#10: ePointEditorName := E_POINT_NAME.HOME_SAFETY; uiPointStorageIndex := UINT#13;
		UINT#11: ePointEditorName := E_POINT_NAME.MAGAZINE_1_DETAIL; uiPointStorageIndex := UINT#14;
		UINT#12: ePointEditorName := E_POINT_NAME.MAGAZINE_2_DETAIL; uiPointStorageIndex := UINT#15;
	ELSE
		ePointEditorName := E_POINT_NAME.NONE;
	END_CASE;

	IF (ePointEditorName <> E_POINT_NAME.NONE) AND (uiPointStorageIndex <> UINT#0) THEN
		GVL_POINT.Points[ePointEditorName] := Persistent_Value.astRetainPoints[uiPointStorageIndex];
		IF (ePointEditorName = E_POINT_NAME.MAGAZINE_1_DETAIL)
		OR (ePointEditorName = E_POINT_NAME.MAGAZINE_2_DETAIL) THEN
			GVL_POINT.Points[ePointEditorName].xConfigured :=
				Persistent_Value.astRetainPoints[uiPointStorageIndex].xConfigured
				AND (Persistent_Value.astRetainPoints[uiPointStorageIndex].MagazineSafeZ <> LREAL#0.0)
				AND (Persistent_Value.astRetainPoints[uiPointStorageIndex].MagazineChangeZ <> LREAL#0.0);
		END_IF;
		IF NOT GVL_POINT.Points[ePointEditorName].xConfigured THEN
			xPointTableReady := FALSE;
		END_IF;
	ELSE
		xPointTableReady := FALSE;
	END_IF;
END_FOR;

// Полнота таблицы остаётся диагностикой редактора. Включение оборудования
// проверяет только собственные точки; HOME_SAFETY отдельно нужен автоциклу.
axMachinePointsReady[1] := GVL_POINT.Points[E_POINT_NAME.MACHINE_1_ABOVE].xConfigured
	AND GVL_POINT.Points[E_POINT_NAME.MACHINE_1_CHUCK_APROACH].xConfigured
	AND GVL_POINT.Points[E_POINT_NAME.MACHINE_1_CHUCK_POSITION].xConfigured;
axMachinePointsReady[2] := GVL_POINT.Points[E_POINT_NAME.MACHINE_2_ABOVE].xConfigured
	AND GVL_POINT.Points[E_POINT_NAME.MACHINE_2_CHUCK_APROACH].xConfigured
	AND GVL_POINT.Points[E_POINT_NAME.MACHINE_2_CHUCK_POSITION].xConfigured;
axMachinePointsReady[3] := GVL_POINT.Points[E_POINT_NAME.MACHINE_3_ABOVE].xConfigured
	AND GVL_POINT.Points[E_POINT_NAME.MACHINE_3_CHUCK_APROACH].xConfigured
	AND GVL_POINT.Points[E_POINT_NAME.MACHINE_3_CHUCK_POSITION].xConfigured;
axMagazinePointsReady[1] := GVL_POINT.Points[E_POINT_NAME.MAGAZINE_1_DETAIL].xConfigured;
axMagazinePointsReady[2] := GVL_POINT.Points[E_POINT_NAME.MAGAZINE_2_DETAIL].xConfigured;

(* ---- PLC_PRG.st ---- *)
PROGRAM PLC_PRG
VAR
    xHmiTablesInitialized : BOOL;
    axTwinStoreChanged : ARRAY [1..2] OF BOOL; // Изменения владельцев, без обхода слотов при публикации
    xGeometryWaitWarningActive : BOOL;
    STATISTIC_MAIN : FB_STATISTIC; // Сбор каждый скан, расчёт раз в 100 мс
	GEOMETRY : ARRAY [1..2] OF FB_GEOMETRY_CONTROL;
	GEOMETRY_SIM : ARRAY [1..2] OF FB_GEOMETRY_CONTROL_SIMULATION;
	xGeometryInitialized : BOOL;
	xGeometryEnvironmentChanged : BOOL;
	eGeometryPreviousEnvironment : E_CELL_TEST_ENVIRONMENT;
	uiGeometry : UINT;
	uiGeometryMachine : UINT;
	uiGeometryDi : UINT;
	udiGeometryRequest : UDINT;
	stGeometryRequest : ST_GEOMETRY_REQUEST;
	stGeometryConfig : ST_GEOMETRY_CONFIG;
	stGeometryCall : ST_GEOMETRY_CALL;
	stGeometryEmptyCall : ST_GEOMETRY_CALL;
	xGeometryConfigValid : BOOL;
	xGeometryDriveAlarm : BOOL;
	xGeometryDriveRunning : BOOL;
	xGeometryPartAtEnd : BOOL;
	stGeometrySignals : ST_GEOMETRY_SIGNALS;
	xGeometryRequestFresh : BOOL;
	xGeometryStopAttempt : BOOL;
	eGeometryPlace : E_POINT_NAME;
	eGeometrySafe : E_POINT_NAME;
	eGeometryChange : E_POINT_NAME;
    // Диагностика физического I/O: один владелец подмен и FIFO на 100 событий.
    axIoRawDi : ARRAY [1..84] OF BOOL;
    axIoUsedDi : ARRAY [1..84] OF BOOL;
    axIoForced : ARRAY [1..84] OF BOOL;
    axIoForceValue : ARRAY [1..84] OF BOOL;
    axIoDoForced : ARRAY [1..50] OF BOOL;
    xIoSnapshotPublishing : BOOL;
    axIoDoForceValue : ARRAY [1..50] OF BOOL;
    axIoDoInhibited : ARRAY [1..50] OF BOOL;
    axIoDoAllowed : ARRAY [1..50] OF BOOL;
    axIoDoOnAllowed : ARRAY [1..50] OF BOOL;
    axIoGripperBase : ARRAY [1..3] OF BOOL;
    axIoAutoDo : ARRAY [1..50] OF BOOL;
    axIoMagazineInvalidated : ARRAY [1..2] OF BOOL;
    xIoRawSafetyOk : BOOL;
    xIoManualActive : BOOL;
    xIoManualEndedByOperator : BOOL;
    xIoDoRejected : BOOL;
    xIoEmergencyResetRejected : BOOL;
    xIoEmergencyResetRequested : BOOL;
    udiIoEmergencyRequestSeq : UDINT;
    axIoOutput : ARRAY [1..50] OF BOOL;
    axIoPreviousRaw : ARRAY [1..84] OF BOOL;
    axIoPreviousUsed : ARRAY [1..84] OF BOOL;
    axIoPreviousOutput : ARRAY [1..50] OF BOOL;
    astIoEvent : ARRAY [1..100] OF ST_PHYSICAL_IO_EVENT;
    xIoInitialized : BOOL;
    xIoOverrideRejected : BOOL;
    xIoBusy : BOOL;
    uiIoIndex : UINT;
    uiIoWord : UINT;
    uiIoBit : UINT;
    dwIoBit : DWORD;
    udiIoNowMs : UDINT;
    udiIoLastTickMs : UDINT;
    uliIoClockMs : ULINT;
    udiIoHeartbeatSeen : UDINT;
    uliIoLeaseAgeMs : ULINT;
    tonIoOverrideWatchdog : TON;
    udiIoRequestSeq : UDINT;
    uiIoRequestAction : UINT;
    uiIoRequestIndex : UINT;
    xIoRequestValue : BOOL;
	xPhysicalNormal : BOOL;
	xPhysicalWasNormal : BOOL;
	xPhysicalInputEnable : BOOL;
	xPhysicalOutputEnable : BOOL;
	xPhysicalOutputWasEnabled : BOOL;
	uiPhysicalInput : UINT;
	tPhysicalRise : TIME;
	tPhysicalFall : TIME;
	axPhysicalRaw : ARRAY [1..84] OF BOOL;
	axPhysicalFiltered : ARRAY [1..80] OF BOOL;
	axPhysicalButtonArmed : ARRAY [1..80] OF BOOL;
	afbPhysicalInputFilter : ARRAY [1..80] OF FB_DI_FILTER;
	astMachineStatusRaw : ARRAY [1..3] OF ST_MACHINE_IO_STATUS;
	AXIS_X         : FB_AXIS; // Управление осью X
	AXIS_Y         : FB_AXIS; // Управление осью Y
	AXIS_Z         : FB_AXIS; // Управление осью Z
	GROUP_XYZ      : FB_AXIS_GROUP; // Управление группой осей XYZ
	SIMULATION_DYNAMICS : FB_SIMULATION_DYNAMIC_LIMITS; // Транзакционное масштабирование лимитов XYZ между тестами
	MOTION_MANAGER : FB_MOTION_MANAGER; // Менеджер движения по именованным точкам
	MACHINE_1      : FB_MACHINE; // Логика первого станка
	MACHINE_2      : FB_MACHINE; // Логика второго станка
	MACHINE_3      : FB_MACHINE; // Логика третьего станка
	MACHINE_1_SIM  : FB_MACHINE_SIMULATION; // Симуляция первого станка
	MACHINE_2_SIM  : FB_MACHINE_SIMULATION; // Симуляция второго станка
	MACHINE_3_SIM  : FB_MACHINE_SIMULATION; // Симуляция третьего станка
	MACHINE_1_FAULT: FB_MACHINE_FAULT_INJECTOR; // Инъекция обратной связи первого станка
	MACHINE_2_FAULT: FB_MACHINE_FAULT_INJECTOR; // Инъекция обратной связи второго станка
	MACHINE_3_FAULT: FB_MACHINE_FAULT_INJECTOR; // Инъекция обратной связи третьего станка
	TWIN_AXIS_1 : FB_AXIS;
	TWIN_AXIS_2 : FB_AXIS;
	TWIN : ARRAY [1..2] OF FB_TWO_PALLET;
	axTwinMagazineExchangeInProgress : ARRAY [1..2] OF BOOL; // Защёлка фактической смены палет для адресной блокировки магазина
	TWIN_SIM : ARRAY [1..2] OF FB_TWO_PALLET_SIMULATION;
	astTwinCommand : ARRAY [1..2] OF ST_TWO_PALLET_COMMAND;
	axTwinConfigurationChanged : ARRAY [1..2] OF BOOL;
	axTwinExternalCommandRejected : ARRAY [1..2] OF BOOL;
	audiTwinWarningSeen : ARRAY [1..2] OF UDINT;
	audiPartWarningSeen : ARRAY [1..2] OF UDINT;
	astMagazineWarningMerged : ARRAY [1..2] OF ST_WARNING_EVENT;
	uiTwin : UINT;
	uiTwinPallet : UINT;
	uiTwinRobotPalletBefore : UINT; // Смена роли после ручного восстановления снимает прежнюю готовность загрузки
	uiTwinSlot : UINT;
	udiTwinSnapshot : UDINT;
	xTwinStartup : BOOL;
	xTwinSimulationInitialized : BOOL;
	axTwinSimIoOwned : ARRAY [1..2] OF BOOL;
	axTwinSafetyBusy : ARRAY [1..2] OF BOOL;
	axButtonStationInput : ARRAY [1..4] OF BOOL; // Физическая кнопка или виртуальный вход SIMULATION
	axButtonStationEmergencyStopInput : ARRAY [1..4] OF BOOL; // Физический грибок или виртуальный вход SIMULATION
	axTwinRobotStopLatched : ARRAY [1..2] OF BOOL;
	xTwinRobotSwapWindow : BOOL;
	xTwinRobotOperation : BOOL; // Текущая, ожидающая отключения или уже выданная операция магазина
	xTwinOtherLoaded : BOOL;
	xTwinRobotHasBlank : BOOL; // Любая заготовка рабочего банка запрещает автоматический обмен
	xTwinOtherHasBlank : BOOL; // Подтверждённая операторская палета должна содержать заготовку
	xTwinInventoryEditPending : BOOL; // Правка текущего скана отменяет запуск по старому подтверждению
	xTwinAutoSwapEnabled : BOOL;
	axTwinAutoSwapPending : ARRAY [1..2] OF BOOL; // Ожидание смены Finished либо отменяемый ранний запрос
	axMagazineInventoryChanged : ARRAY [1..2] OF BOOL; // Смена/правка только рабочего банка снимает его Finished
	xTwinInventoryCommand : BOOL;
	uiTwinRequestResult : UINT;
	stTwinRequest : ST_TWO_PALLET_REQUEST;
	fbMagazine1    : FB_MAGAZINE; // Первый статичный магазин
	fbMagazine2    : FB_MAGAZINE; // Второй статичный магазин
	ROBOT          : FB_ROBOT; // Координация движений и захвата робота
	stRobotResetDependencies : ST_ROBOT_RESET_DEPENDENCIES; // Внутренний снимок владельцев зависимого Stop
	ROBOT_MODBUS   : FB_ROBOT_MODBUS; // Modbus TCP транспорт внешнего контроллера
	TYPE_CONFIG    : FB_MULTI_TYPE_CONFIG_MANAGER; // Конфигурация типов продукции
	CELL_SAFETY    : FB_CELL_SAFETY; // Дискретный контур безопасности, двери и внешние кнопки
	CELL_MANAGER   : FB_CELL_MANAGER; // Универсальный автоматический цикл для одного-трёх типов
	ALARM_MANAGER  : FB_ALARM_MANAGER; // Журнал аварий и предупреждений
    CONTROLLER_DIAGNOSTICS : FB_CONTROLLER_DIAGNOSTICS;
	fbAlarmHorn : FB_ALARM_HORN; // Импульс на каждую новую аварийную маску
	tonSignalTowerBlink : TON; // Полупериод мигания колонны — 500 мс
	usiSignalTowerMode : USINT; // 1 работа; 2 готова; 3 предупреждение; 4 авария; 5 не готова
	usiSignalTowerPreviousMode : USINT;
	xSignalTowerBlinkOn : BOOL := TRUE;
	uiHmiCommandIndex : UINT;
	udiHmiCommandNowMs : UDINT;
	axHmiCommandConsumed : ARRAY [1..121] OF BOOL;
	axHmiCommandWasHigh : ARRAY [1..121] OF BOOL;
	axHmiInternalPulse : ARRAY [1..121] OF BOOL; // Internal scenario events, consumed next scan
	axHmiCommandPulse : ARRAY [1..121] OF BOOL;
	audiHmiCommandSnapshot : ARRAY [1..121] OF UDINT;
	udiCellSettingSnapshot : UDINT;
	xCellSettingRejected : BOOL;
	uiMachine      : UINT; // Индекс станка при обработке команд HMI
	iDetail        : SINT; // Индекс слота при передаче состояния магазина в HMI
	xRobotHmiPermit: BOOL; // Разрешение ручных команд робота с HMI
	udiCellModeCommandSnapshot : UDINT; // Снимок маркера транзакции текущего скана
	uiCellModeRejectReason : UINT; // Одноцикловая причина отказа для журнала ячейки
	xDrivesReady   : BOOL; // Все оси и группа готовы к движению
	xDrivesPowered : BOOL; // На все три оси фактически подано питание
	xAnyDrivePowered : BOOL; // Хотя бы на одну ось фактически подано питание
	xDrivesOff     : BOOL; // Все силовые части отключены, группа в GroupDisabled
	xPowerTransitionActive : BOOL; // Выполняется последовательность включения или отключения
	xPowerDisableRequest : BOOL; // Единый запрос штатного отключения через группу
	xDriveError    : BOOL; // Активна ошибка хотя бы одной оси или группы
	xAxisDriveError : BOOL; // Активна ошибка одиночной оси; не включает административную ошибку группы
	xGroupError    : BOOL; // Активна ошибка координатной группы
	xMotionBusy    : BOOL; // Хотя бы одна ось ещё выполняет команду
	xGroupMotionBusy : BOOL; // Координатная группа выполняет движение или остановку
	xRobotAutoPowerOff : BOOL; // Автоматическое снятие питания приводов при аварии робота
	xHmiConnectionAlive : BOOL; // Watchdog связи HMI -> PLC
	xManualRecoveryActive : BOOL; // Ограниченное ручное восстановление при общей ошибке
	xHmiRobotActionBaseAllowed : BOOL; // Условия ручного перемещения робота к точке
	xHmiRobotPointTargetAllowed : BOOL; // Люк соответствующего станка открыт для входной точки
	xHmiRobotPointAllowed : BOOL; // Полное разрешение выбранной ручной точки
	eHmiRobotStatusAction : E_ROBOT_ACTION; // Действие для отображения xAllowed/reason
	eHmiRobotStatusPoint : E_POINT_NAME; // Точка для отображения xAllowed/reason
	xHmiRobotStatusPointTargetAllowed : BOOL; // Безопасность выбранной HMI-точки
	xHmiRobotStatusPointAllowed : BOOL; // Полное разрешение выбранной HMI-точки
	xHmiGripperActionBaseAllowed : BOOL; // Условия ручного действия захвата независимо от Motion-слоя
	xHmiRobotActionAllowed : BOOL;
	xHmiRobotActionAttempt : BOOL;
	rtHmiRobotAction : R_TRIG;
	udiLastHmiHeartbeat : UDINT; // Последний принятый heartbeat HMI
	tonHmiWatchdog : TON; // Таймаут HMI heartbeat
	udiLastMobileMotionHeartbeat : UDINT; // Последний heartbeat мобильной аренды
	tonMobileMotionWatchdog : TON; // Таймаут gateway/телефон -> PLC для мобильного движения
	rtMobileMotionStart : R_TRIG; // Фронт новой мобильной аренды
	xMobileMotionLeaseActive : BOOL; // PLC защёлкнул мобильного владельца до полного останова
	xMobileMotionConnectionAlive : BOOL; // Мобильный heartbeat обновляется
	xMobileMotionStopRequest : BOOL; // Независимый запрос контролируемой остановки оси
	rMobileMotionSpeedLimitPercent : REAL := 0.1; // Защёлкнутый глобальный лимит телефона
	rRobotManualEffectiveSpeedPercent : REAL := 0.1; // Итоговый override после PLC-ограничения
	uiManualAxisOwner : UINT; // Единственная ось-владелец текущей команды HMI
	uiManualAxisRequest : UINT; // Ось, запросившая новую ручную команду в текущем цикле
	axManualAxisBaseAllowed : ARRAY [1..3] OF BOOL;
	axManualAxisCommandRejected : ARRAY [1..3] OF BOOL;
	artManualAxisReject : ARRAY [1..3] OF R_TRIG;
	artHmiAxisHome : ARRAY [1..3] OF R_TRIG; // Фронты импульсных Home-команд HMI
	artHmiAxisMoveAbsolute : ARRAY [1..3] OF R_TRIG; // Фронты абсолютных команд HMI
	artHmiAxisMoveRelative : ARRAY [1..3] OF R_TRIG; // Фронты шаговых команд HMI
	axHmiAxisHomePulse : ARRAY [1..3] OF BOOL;
	axHmiAxisMoveAbsolutePulse : ARRAY [1..3] OF BOOL;
	axHmiAxisMoveRelativePulse : ARRAY [1..3] OF BOOL;
	alrRobotManualRatedVelocity : ARRAY [1..3] OF LREAL; // Фактические 100% из AXIS_REF_SM3
	alrRobotRatedAcceleration : ARRAY [1..3] OF LREAL; // Максимальное ускорение из AXIS_REF_SM3
	alrRobotRatedDeceleration : ARRAY [1..3] OF LREAL; // Максимальное замедление из AXIS_REF_SM3
	alrRobotRatedJerk : ARRAY [1..3] OF LREAL; // Максимальный jerk из AXIS_REF_SM3
	axRobotSoftwareLimitsEnabled : ARRAY [1..3] OF BOOL; // Фактическое включение software limits в AXIS_REF_SM3
	alrRobotSoftwareMinPosition : ARRAY [1..3] OF LREAL; // Отрицательный software limit SoftMotion
	alrRobotSoftwareMaxPosition : ARRAY [1..3] OF LREAL; // Положительный software limit SoftMotion
	alrRobotJogVelocity : ARRAY [1..3] OF LREAL; // Скорость одиночной оси с учётом общего коэффициента
	xHmiDrivesEnableAccepted : BOOL; // Авторитетное решение RunMotion по команде включения
	xHmiDrivesDisableAccepted : BOOL; // Авторитетное решение RunMotion по команде отключения
	xHmiResetAccepted : BOOL; // Авторитетное решение RunMotion по команде сброса
	xHmiStopAccepted : BOOL; // Авторитетное решение RunMotion по команде остановки
	xRobotMotionCommandActive : BOOL; // Принятая команда, включая проверку точки и освобождение
	xRobotProgramStopRequest : BOOL; // Штатная остановка группового движения по запросу автоматики
	xMotionResetRequest : BOOL; // Общий запрос последовательного сброса группы и осей
	xGroupResetPulse : BOOL; // Импульс MC_GroupReset; он также сбрасывает оси группы
	xAxisResetPulse : BOOL; // Последующая очистка локальных защёлок FB_AXIS
	xMotionResetBusy : BOOL; // Последовательность сброса Motion-слоя активна
	rtMotionReset : R_TRIG; // Фронт единого запроса сброса Motion-слоя
	eMotionResetState : E_MOTION_RESET_STATE := E_MOTION_RESET_STATE.IDLE;
	xAlarmResetRequired : BOOL; // Хотя бы один владелец общей команды находится в аварии
	xAlarmResetAllowed : BOOL; // Все активные владельцы аварий готовы принять общий сброс
	stRobotHmiCommand : ST_ROBOT_COMMAND; // Команда робота с учётом оперативной остановки HMI
	stSelectedMagazineCommand : ST_ROBOT_COMMAND; // Единственная команда двух магазинов роботу
	stMagazinePointCommand : ST_ROBOT_COMMAND; // Команда, по которой рассчитывается временная точка
	eMagazineBasePoint : E_POINT_NAME; // База выбранного магазина
	uiMagazine : UINT; // Индекс магазина 1..2
	auiMagazineEditSlot : ARRAY [1..2] OF UINT; // Новый контракт с fallback на legacy-команду первого магазина
	astMachineFaultRequest : ARRAY [1..3] OF ST_MACHINE_FAULT_REQUEST; // Запросы ошибок станков
	astAxisFaultRequest    : ARRAY [1..3] OF ST_AXIS_FAULT_REQUEST; // Запросы ошибок осей
	stAxisGroupFaultRequest: ST_AXIS_GROUP_FAULT_REQUEST; // Запрос ошибки группы XYZ
	stRobotFaultRequest    : ST_ROBOT_FAULT_REQUEST; // Запросы ошибок робота и точки
	astMagazineFaultRequest : ARRAY [1..2] OF ST_MAGAZINE_FAULT_REQUEST; // Диагностика двух магазинов
	stCellFaultRequest     : ST_CELL_FAULT_REQUEST; // Запрос локальной ошибки менеджера ячейки
	stSafetyFaultRequest   : ST_CELL_SAFETY_FAULT_REQUEST; // Независимые инъекции дискретной безопасности
	astAlarmSource : ARRAY [1..22] OF ST_ALARM_SOURCE_DATA; // Старые коды сохранены; диагностика MC522 добавлена в конец.
	astAdditionalCellWarning : ARRAY [1..2] OF ST_WARNING_EVENT; // 1: конфигуратор, 2: общие предупреждения ГК
	uiPointEditorIndex : UINT; // Компактный индекс фиксированной точки редактора 1..14
	uiPointEditorGeometryStation : UINT; // 0 прежняя точка, 1/2 база ГК
	uiPointStorageIndex : UINT; // Индекс в совместимом Persistent-массиве 1..15
	ePointEditorName : E_POINT_NAME; // Фактический enum выбранной инженерной точки
	xPointTableReady : BOOL; // Все 12 базовых точек подтверждены редактором
	axMachinePointsReady : ARRAY [1..3] OF BOOL; // Три рабочие точки каждого станка
	axMagazinePointsReady : ARRAY [1..2] OF BOOL; // Полная калибровка выбранного метода каждого магазина
	astMagazineFrame : ARRAY [1..2] OF ST_MAGAZINE_FRAME;
	uiCalibrationMagazine : UINT;
	eCalibrationOrigin : E_POINT_NAME;
	eCalibrationPointB : E_POINT_NAME;
	eCalibrationPointC : E_POINT_NAME;
	uiPointEditorMagazine : UINT;
	uiPointEditorReference : UINT;
	uiCalibrationSettingMagazine : UINT;
	xMagazineCalibrationEditAllowed : ARRAY [1..2] OF BOOL;
	stMagazineReferenceDraft : ST_POINT;
	xCellPointsReady : BOOL; // HOME_SAFETY и точки только включённого оборудования
	xPointEditorBaseAllowed : BOOL; // Общие безопасные условия Capture/Save
	xPointEditorAllHomed : BOOL; // Все оси XYZ прошли Home
	xPointEditorRequestValid : BOOL; // Индекс и код новой транзакции распознаны
	xPointEditorDraftValid : BOOL; // XYZ и скорость черновика прошли проверку
	xPointEditorMagazinePoint : BOOL; // Выбрана базовая точка магазина 1 или 2
	xPointEditorGeometrySave : BOOL; // SAVE базы ГК не зависит от технологических блокировок
	udiLastPointEditorCommandSeq : UDINT; // Последняя обработанная транзакция редактора
	xPointCheckRequest : BOOL;
	xPointCheckActive : BOOL;
	xPointCheckStopping : BOOL;
	xPointCheckSeenBusy : BOOL;
	xPointCheckSeenDone : BOOL; // Терминальный ответ Motion хранится до фактического останова
	xPointCheckStopRequest : BOOL;
	xPointCheckConnectionAlive : BOOL;
	udiLastPointCheckHeartbeat : UDINT;
	tonPointCheckWatchdog : TON;
	tonPointCheckStart : TON;
	ePointCheckName : E_POINT_NAME;
	uiPointCheckLoop : UINT;
	uiPointCheckMachine : UINT;
	uiPointCheckReason : UINT;
	stPointCheckCandidate : ST_POINT;
	rPointCheckLatchedSpeed : REAL;
	lrGroupVelocityOverride : LREAL;
	xRobotInterfaceReady : BOOL; // Готовность применённого интерфейса робота
	lrRobotActualX : LREAL; // Координаты выбранного источника управления
	lrRobotActualY : LREAL;
	lrRobotActualZ : LREAL;
	xModeCommonSafe : BOOL; // Общие условия изменения источника управления
	xAllMachinesIdle : BOOL;
	rtRobotModeApply : R_TRIG;
	rtModbusSettingsApply : R_TRIG;
	xModbusHmiInitialized : BOOL;
	uiRobotInterfaceWarningCode : UINT;
	uiRobotManualMagazineIndex : UINT;
	uiRobotManualMagazineRow : UINT;
	uiRobotManualMagazineColumn : UINT;
	rtTestEnvironmentApply : R_TRIG;
	rtTestSpeedProfileApply : R_TRIG;
	rtTestScenarioApply : R_TRIG;
	xTestInitializePulse : BOOL;
	xTestAbortActive : BOOL; // Тестовая отмена действует только в виртуальной среде
	xTestStable : BOOL;
	xTestScenarioValid : BOOL;
	uiTestIndex : UINT;
	uiTestMagazine : UINT;
	uiTestFaultOwnerCount : UINT;
	uiTestSlotCount : UINT;
	uiTestPallet : UINT;
	uiTestOtherPallet : UINT;
	uiTestType : UINT;
	xTestTypeHasMachine : BOOL;
	xTestTypeHasSlot : BOOL;
	udiTestGeometryProduced : UDINT;
	xTestGeometrySettingsSaved : BOOL;
	xTestSavedGeometryAuto : BOOL;
	xTestSavedGeometryWait : BOOL;
	stTestEmptyGeometryMemory : ST_GEOMETRY_MEMORY;
	stTestEmptyGeometryCall : ST_GEOMETRY_CALL;
	adwTestMagazineFaultMask : ARRAY [1..2] OF DWORD;
	xApplicationStartupInitialized : BOOL; // Однократная инициализация безопасных настроек после старта/Online Change
END_VAR

VAR CONSTANT
	WRN_HMI_MANUAL_REJECTED : UINT := 12; // PLC отклонил команду расширенного ручного управления
	WRN_ROBOT_MODE_REJECTED : UINT := 13; // PLC отклонил переключение источника управления
	WRN_MODBUS_SETTINGS_REJECTED : UINT := 14; // PLC отклонил применение параметров соединения
	WRN_POINT_EDIT_REJECTED : UINT := 15; // PLC отклонил Capture/Save/Invalidate инженерной точки
	WRN_POINT_CHECK_REJECTED : UINT := 16; // Проверка точки отклонена
	WRN_POINT_CHECK_INTERRUPTED : UINT := 17; // Проверка остановлена потерей связи/разрешений
	aePointCheckNames : ARRAY [1..18] OF E_POINT_NAME := [
		E_POINT_NAME.MACHINE_1_ABOVE, E_POINT_NAME.MACHINE_1_CHUCK_APROACH, E_POINT_NAME.MACHINE_1_CHUCK_POSITION,
		E_POINT_NAME.MACHINE_2_ABOVE, E_POINT_NAME.MACHINE_2_CHUCK_APROACH, E_POINT_NAME.MACHINE_2_CHUCK_POSITION,
		E_POINT_NAME.MACHINE_3_ABOVE, E_POINT_NAME.MACHINE_3_CHUCK_APROACH, E_POINT_NAME.MACHINE_3_CHUCK_POSITION,
		E_POINT_NAME.HOME_SAFETY, E_POINT_NAME.MAGAZINE_1_DETAIL, E_POINT_NAME.MAGAZINE_2_DETAIL,
		E_POINT_NAME.GEOMETRY_1_PLACE, E_POINT_NAME.GEOMETRY_2_PLACE,
		E_POINT_NAME.MAGAZINE_1_AXIS_X, E_POINT_NAME.MAGAZINE_1_AXIS_Y,
		E_POINT_NAME.MAGAZINE_2_AXIS_X, E_POINT_NAME.MAGAZINE_2_AXIS_Y];
	alrRobotManualFallbackVelocity : ARRAY [1..3] OF LREAL := [1000.0, 1000.0, 1000.0]; // Резерв, если привод не публикует динамический предел
	alrRobotManualAcceleration : ARRAY [1..3] OF LREAL := [1000.0, 1000.0, 1000.0]; // Резерв ускорения, если привод не публикует предел
	alrRobotManualDeceleration : ARRAY [1..3] OF LREAL := [1000.0, 1000.0, 1000.0]; // Резерв замедления, если привод не публикует предел
	alrRobotManualJerk : ARRAY [1..3] OF LREAL := [10000.0, 10000.0, 10000.0]; // Резерв jerk, если привод не публикует предел
END_VAR

// --- BEGIN IMPLEMENTATION ---

SetApplicationDefaults();
ReadHmiCommands();
ReadHmiInputs();
ReadIoEmergencyStop();
ReadPhysicalInputs();
RunSafety();
ResetIoEmergencyStop();
RunMotion();
RunRobotModbus();
RunTestControl();
RunMagazineCalibration();
RunTwoPallet();
RunGeometryControl();
RunCellControl();
RunMachines();
RunMagazine();
RunTwoPalletAxis();
RunRobot();
RunStatistics();
RunAlarms();
RunSignalTower();
WritePhysicalOutputs();
RecordIoDiagnostics();
PublishGeometryControl();
PublishHmi();

(* ---- PLC_PRG.WritePhysicalOutputs.st ---- *)
METHOD PRIVATE WritePhysicalOutputs

// --- BEGIN IMPLEMENTATION ---

// Единственная страница назначения выходов. Выполняется после всех владельцев команд.
// Не публикуем команды симулятора на железо при смене среды в текущем скане.
xPhysicalOutputEnable := GVL_PHYSICAL_IO.xNormalActive
	AND (GVL_CELL_SETTINGS.eTestEnvironment = E_CELL_TEST_ENVIRONMENT.NORMAL);
IF xPhysicalOutputEnable THEN
	FOR uiMachine := 1 TO 3 DO
		IF GVL_MACHINE.Command[uiMachine].stIo.xCloseDoor
		AND NOT GVL_MACHINE.Command[uiMachine].stIo.xOpenDoor THEN
			GVL_PHYSICAL_IO.axMachineHatchClose[uiMachine] := TRUE;
		ELSIF GVL_MACHINE.Command[uiMachine].stIo.xOpenDoor
		AND NOT GVL_MACHINE.Command[uiMachine].stIo.xCloseDoor THEN
			GVL_PHYSICAL_IO.axMachineHatchClose[uiMachine] := FALSE;
		ELSIF NOT xPhysicalOutputWasEnabled THEN
			GVL_PHYSICAL_IO.axMachineHatchClose[uiMachine] := GVL_MACHINE.astPhysicalInput[uiMachine].xDoorClosed;
		END_IF;
	END_FOR;
	IF NOT GVL_HMI.xModbusMode AND GVL_PHYSICAL_IO.stGripperCommand.xExecute THEN
		CASE GVL_PHYSICAL_IO.stGripperCommand.eAction OF
			E_ROBOT_ACTION.UNCLAMP_1: axIoGripperBase[1] := TRUE;
			E_ROBOT_ACTION.CLAMP_1: axIoGripperBase[1] := FALSE;
			E_ROBOT_ACTION.UNCLAMP_2: axIoGripperBase[2] := TRUE;
			E_ROBOT_ACTION.CLAMP_2: axIoGripperBase[2] := FALSE;
			E_ROBOT_ACTION.ROTATE_TO_BLANK: axIoGripperBase[3] := FALSE;
			E_ROBOT_ACTION.ROTATE_TO_DETAIL: axIoGripperBase[3] := TRUE;
		END_CASE;
	END_IF;
END_IF;
// Внешний SC-500 остаётся единственным владельцем захватов в Modbus.
IF NOT xPhysicalOutputEnable OR GVL_HMI.xModbusMode THEN
	axIoGripperBase[1] := FALSE;
	axIoGripperBase[2] := FALSE;
	axIoGripperBase[3] := FALSE;
END_IF;
GVL_PHYSICAL_IO.xDoGripper1Open := axIoGripperBase[1];
GVL_PHYSICAL_IO.xDoGripper2Open := axIoGripperBase[2];
GVL_PHYSICAL_IO.xDoRotateToDetail := axIoGripperBase[3];

GVL_PHYSICAL_IO.xDoMachine1HatchClosed := xPhysicalOutputEnable AND GVL_PHYSICAL_IO.axMachineHatchClose[1];
GVL_PHYSICAL_IO.xDoMachine1HatchUnLock := xPhysicalOutputEnable AND GVL_MACHINE.Command[1].stIo.xHatchUnLock;
GVL_PHYSICAL_IO.xDoMachine1ClampChuck := xPhysicalOutputEnable AND GVL_MACHINE.Command[1].stIo.xClampChuck AND NOT GVL_MACHINE.Command[1].stIo.xUnclampChuck;
GVL_PHYSICAL_IO.xDoMachine1UnclampChuck := xPhysicalOutputEnable AND GVL_MACHINE.Command[1].stIo.xUnclampChuck AND NOT GVL_MACHINE.Command[1].stIo.xClampChuck;
GVL_PHYSICAL_IO.xDoMachine1StartCycle := xPhysicalOutputEnable AND GVL_MACHINE.Command[1].stIo.xStartCycle;
GVL_PHYSICAL_IO.xDoMachine2HatchClosed := xPhysicalOutputEnable AND GVL_PHYSICAL_IO.axMachineHatchClose[2];
GVL_PHYSICAL_IO.xDoMachine2HatchUnLock := xPhysicalOutputEnable AND GVL_MACHINE.Command[2].stIo.xHatchUnLock;
GVL_PHYSICAL_IO.xDoMachine2ClampChuck := xPhysicalOutputEnable AND GVL_MACHINE.Command[2].stIo.xClampChuck AND NOT GVL_MACHINE.Command[2].stIo.xUnclampChuck;
GVL_PHYSICAL_IO.xDoMachine2UnclampChuck := xPhysicalOutputEnable AND GVL_MACHINE.Command[2].stIo.xUnclampChuck AND NOT GVL_MACHINE.Command[2].stIo.xClampChuck;
GVL_PHYSICAL_IO.xDoMachine2StartCycle := xPhysicalOutputEnable AND GVL_MACHINE.Command[2].stIo.xStartCycle;
GVL_PHYSICAL_IO.xDoMachine3HatchClosed := xPhysicalOutputEnable AND GVL_PHYSICAL_IO.axMachineHatchClose[3];
GVL_PHYSICAL_IO.xDoMachine3HatchUnLock := xPhysicalOutputEnable AND GVL_MACHINE.Command[3].stIo.xHatchUnLock;
GVL_PHYSICAL_IO.xDoMachine3ClampChuck := xPhysicalOutputEnable AND GVL_MACHINE.Command[3].stIo.xClampChuck AND NOT GVL_MACHINE.Command[3].stIo.xUnclampChuck;
GVL_PHYSICAL_IO.xDoMachine3UnclampChuck := xPhysicalOutputEnable AND GVL_MACHINE.Command[3].stIo.xUnclampChuck AND NOT GVL_MACHINE.Command[3].stIo.xClampChuck;
GVL_PHYSICAL_IO.xDoMachine3StartCycle := xPhysicalOutputEnable AND GVL_MACHINE.Command[3].stIo.xStartCycle;
GVL_PHYSICAL_IO.xDoDoor1Unlock := xPhysicalOutputEnable AND GVL_CELL_SAFETY_IO.axDoorUnlockOutput[1];
GVL_PHYSICAL_IO.xDoDoor2Unlock := xPhysicalOutputEnable AND GVL_CELL_SAFETY_IO.axDoorUnlockOutput[2];
GVL_PHYSICAL_IO.xDoDoor3Unlock := xPhysicalOutputEnable AND GVL_CELL_SAFETY_IO.axDoorUnlockOutput[3];
GVL_PHYSICAL_IO.xDoDoor4Unlock := xPhysicalOutputEnable AND GVL_CELL_SAFETY_IO.axDoorUnlockOutput[4];
GVL_PHYSICAL_IO.xDoSafetyRelayReset := xPhysicalOutputEnable AND GVL_CELL_SAFETY_IO.xSafetyRelayResetOutput;
GVL_PHYSICAL_IO.xDoSignalTowerGreenOutput := xPhysicalOutputEnable AND GVL_CELL_SAFETY_IO.xSignalTowerGreenOutput;
GVL_PHYSICAL_IO.xDoSignalTowerAmberOutput := xPhysicalOutputEnable AND GVL_CELL_SAFETY_IO.xSignalTowerAmberOutput;
GVL_PHYSICAL_IO.xDoSignalTowerRedOutput := xPhysicalOutputEnable AND GVL_CELL_SAFETY_IO.xSignalTowerRedOutput;
GVL_PHYSICAL_IO.xDoDoor1ButtonLamp := xPhysicalOutputEnable AND GVL_CELL_SAFETY_IO.axDoorButtonLampOutput[1];
GVL_PHYSICAL_IO.xDoDoor2ButtonLamp := xPhysicalOutputEnable AND GVL_CELL_SAFETY_IO.axDoorButtonLampOutput[2];
GVL_PHYSICAL_IO.xDoDoor3ButtonLamp := xPhysicalOutputEnable AND GVL_CELL_SAFETY_IO.axDoorButtonLampOutput[3];
GVL_PHYSICAL_IO.xDoDoor4ButtonLamp := xPhysicalOutputEnable AND GVL_CELL_SAFETY_IO.axDoorButtonLampOutput[4];
GVL_PHYSICAL_IO.xDoMagazine1LockIn := xPhysicalOutputEnable AND (GVL_TWO_PALLET.uiMode = UINT#1) AND GVL_TWO_PALLET.astOutput[1].xLockIn AND NOT GVL_TWO_PALLET.astOutput[1].xLockOut;
GVL_PHYSICAL_IO.xDoMagazine1LockOut := xPhysicalOutputEnable AND (GVL_TWO_PALLET.uiMode = UINT#1) AND GVL_TWO_PALLET.astOutput[1].xLockOut AND NOT GVL_TWO_PALLET.astOutput[1].xLockIn;
GVL_PHYSICAL_IO.xDoMagazine1StopIn := xPhysicalOutputEnable AND (GVL_TWO_PALLET.uiMode = UINT#1) AND GVL_TWO_PALLET.astOutput[1].xStopIn AND NOT GVL_TWO_PALLET.astOutput[1].xStopOut;
GVL_PHYSICAL_IO.xDoMagazine1StopOut := xPhysicalOutputEnable AND (GVL_TWO_PALLET.uiMode = UINT#1) AND GVL_TWO_PALLET.astOutput[1].xStopOut AND NOT GVL_TWO_PALLET.astOutput[1].xStopIn;
GVL_PHYSICAL_IO.xDoMagazine1LiftUp := xPhysicalOutputEnable AND (GVL_TWO_PALLET.uiMode = UINT#1) AND GVL_TWO_PALLET.astOutput[1].xLiftUp AND NOT GVL_TWO_PALLET.astOutput[1].xLiftDown;
GVL_PHYSICAL_IO.xDoMagazine1LiftDown := xPhysicalOutputEnable AND (GVL_TWO_PALLET.uiMode = UINT#1) AND GVL_TWO_PALLET.astOutput[1].xLiftDown AND NOT GVL_TWO_PALLET.astOutput[1].xLiftUp;
GVL_PHYSICAL_IO.xDoMagazine2LockIn := xPhysicalOutputEnable AND (GVL_TWO_PALLET.uiMode = UINT#1) AND GVL_TWO_PALLET.astOutput[2].xLockIn AND NOT GVL_TWO_PALLET.astOutput[2].xLockOut;
GVL_PHYSICAL_IO.xDoMagazine2LockOut := xPhysicalOutputEnable AND (GVL_TWO_PALLET.uiMode = UINT#1) AND GVL_TWO_PALLET.astOutput[2].xLockOut AND NOT GVL_TWO_PALLET.astOutput[2].xLockIn;
GVL_PHYSICAL_IO.xDoMagazine2StopIn := xPhysicalOutputEnable AND (GVL_TWO_PALLET.uiMode = UINT#1) AND GVL_TWO_PALLET.astOutput[2].xStopIn AND NOT GVL_TWO_PALLET.astOutput[2].xStopOut;
GVL_PHYSICAL_IO.xDoMagazine2StopOut := xPhysicalOutputEnable AND (GVL_TWO_PALLET.uiMode = UINT#1) AND GVL_TWO_PALLET.astOutput[2].xStopOut AND NOT GVL_TWO_PALLET.astOutput[2].xStopIn;
GVL_PHYSICAL_IO.xDoMagazine2LiftUp := xPhysicalOutputEnable AND (GVL_TWO_PALLET.uiMode = UINT#1) AND GVL_TWO_PALLET.astOutput[2].xLiftUp AND NOT GVL_TWO_PALLET.astOutput[2].xLiftDown;
GVL_PHYSICAL_IO.xDoMagazine2LiftDown := xPhysicalOutputEnable AND (GVL_TWO_PALLET.uiMode = UINT#1) AND GVL_TWO_PALLET.astOutput[2].xLiftDown AND NOT GVL_TWO_PALLET.astOutput[2].xLiftUp;

GVL_PHYSICAL_IO.xDoCellAlarmHorn := xPhysicalOutputEnable AND GVL_CELL_SAFETY_IO.xAlarmHornOutput;
GVL_PHYSICAL_IO.xDoGk1DriveRun := xPhysicalOutputEnable AND GEOMETRY[1].xRunOutput;
GVL_PHYSICAL_IO.xDoGk1DriveReset := xPhysicalOutputEnable AND GEOMETRY[1].xResetOutput;

GVL_PHYSICAL_IO.xDoGk2DriveRun := xPhysicalOutputEnable AND GEOMETRY[2].xRunOutput;
GVL_PHYSICAL_IO.xDoGk2DriveReset := xPhysicalOutputEnable AND GEOMETRY[2].xResetOutput;

ApplyIoOutputOverrides();

xPhysicalOutputWasEnabled := xPhysicalOutputEnable;

(* ---- STATISTIC.st ---- *)
PROGRAM STATISTIC
VAR
END_VAR

// --- BEGIN IMPLEMENTATION ---

// Совместимость со старой Task Configuration: программа больше не пишет данные.
// Сбор и расчёт перенесены в PLC_PRG.RunStatistics, единственный владелец — MainTask.
// После импорта удалить вызов STATISTIC и отдельную StatisticTask в CODESYS.
